REGION Network 18: MUTE 2
   RUNG wire#powerrail
      #Mute_LG_2_DB("I_S_Time_extension (TE)" := wire#w1, I_S_Material_selection_1 := wire#w2, "########## BASIC_INPUTS ##########" :=, I_S_ESPE_Channel_1 := #Light_Guard_Tuned, I_S_ESPE_Channel_2 := #Light_Guard_Tuned, "I_S_PLC_request (MR)" := #MR_2, I_S_Reset := #ACK, "I_S_Override hold-to-run-device" := #Bypass."Light Guards CX201 - CH1", I_S_first_logic_cycle := "FirstScan", I_S_Disc_Time_MR_and_TE :=, "########## MATERIAL_SELECTION_INPUTS ##########" :=, I_S_Material_selection_2 := #Material_Selection_2, I_S_Material_selection_3 :=, I_S_Material_selection_4 :=, "########## MATERIAL_TOLERANCE_LENGTH in mm ##########" :=, "I_S_Material_tolerance_length_Material_1-4" :=, "########## MAX_DISTANCE_MATERIAL_ESPE in mm ##########" :=, I_S_Max_distance_Material_to_ESPE := 200, "########## MATERIAL_LENGH_1-4 in mm ##########" :=, I_S_Material_length_Material_1 := 1000, I_S_Material_length_Material_2 := 800, I_S_Material_length_Material_3 :=, I_S_Material_length_Material_4 :=, "########## MATERIAL_SPEED_1-4 in mm/s ##########" :=, I_S_Material_speed_Material_1 := 167, I_S_Material_speed_Material_2 := 167, I_S_Material_speed_Material_3 :=, I_S_Material_speed_Material_4 :=, "########## BASIC_OUTPUTS ##########" =>, Q_Safety_release_1 =>, Q_Safety_release_2 =>, Q_SEE_Status =>, Q_Override_Status =>, Q_Reset_required =>, Q_Sequence_OK =>, "########## ERRORS ##########" =>, Error =>)
   END_RUNG
   RUNG wire#powerrail
      I_Contact( #MR_2 )
   END_RUNG wire#w1
   RUNG wire#powerrail
      I_Contact( #Material_Selection_2 )
   END_RUNG wire#w2
   // the same network as SCL:
   #Mute_LG_2_DB(I_S_ESPE_Channel_1 := #Light_Guard_Tuned,   // "SICK Safe Entry Exit HW PLC V02"
                 I_S_ESPE_Channel_2 := #Light_Guard_Tuned,
                 "I_S_PLC_request (MR)" := #MR_2,
                 "I_S_Time_extension (TE)" := NOT #MR_2,
                 I_S_Reset := #ACK,
                 "I_S_Override hold-to-run-device" := #Bypass."Light Guards CX201 - CH1",
                 I_S_first_logic_cycle := "FirstScan",
                 I_S_Material_selection_1 := NOT #Material_Selection_2,
                 I_S_Material_selection_2 := #Material_Selection_2,
                 I_S_Max_distance_Material_to_ESPE := 200,
                 I_S_Material_length_Material_1 := 1000,
                 I_S_Material_length_Material_2 := 800,
                 I_S_Material_speed_Material_1 := 167,
                 I_S_Material_speed_Material_2 := 167);
END_REGION

REGION Network 19: Gate 1 Sensor
   RUNG wire#powerrail
      #Gate_1_DB.ESTOP1(E_STOP := wire#w1, ACK_NEC :=, ACK := #ACK, TIME_DEL :=, Q =>, Q_DELAY =>, ACK_REQ =>, DIAG =>)
   END_RUNG
   RUNG wire#powerrail
      Contact( #Gate_1 )
   END_RUNG wire#w1
   RUNG wire#powerrail
      Contact( #Bypass.Gate_1 )
   END_RUNG wire#w1
   // the same network as SCL:
   #Gate_1_DB(E_STOP := #Gate_1 OR #Bypass.Gate_1, ACK := #ACK);   // ESTOP1
END_REGION

REGION Network 20: Gate 2 Sensor
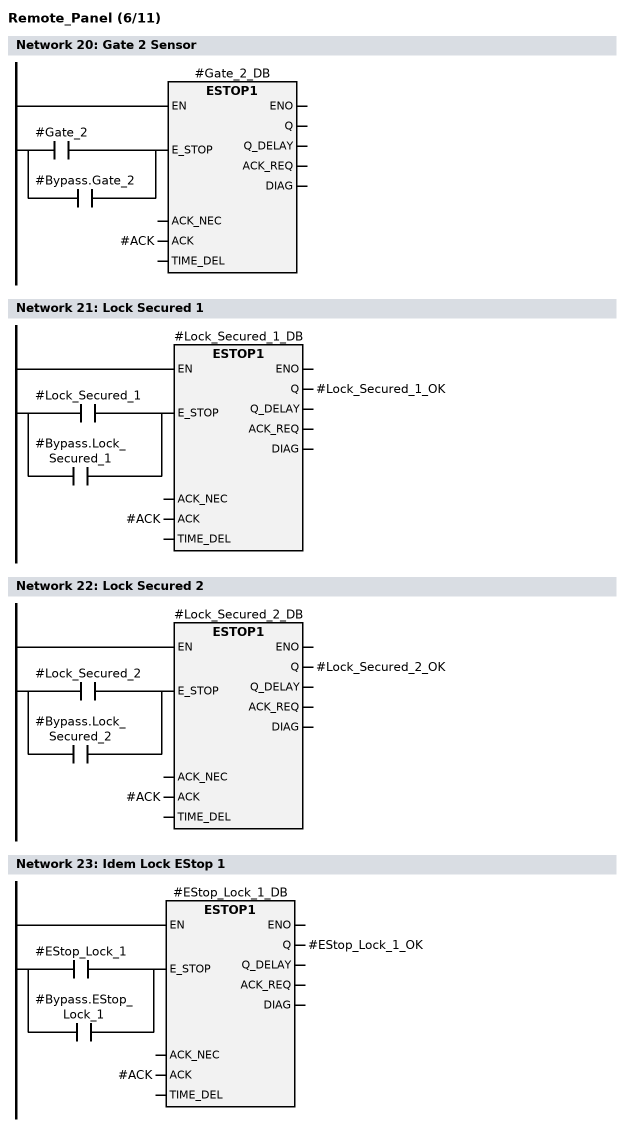
   RUNG wire#powerrail
      #Gate_2_DB.ESTOP1(E_STOP := wire#w1, ACK_NEC :=, ACK := #ACK, TIME_DEL :=, Q =>, Q_DELAY =>, ACK_REQ =>, DIAG =>)
   END_RUNG
   RUNG wire#powerrail
      Contact( #Gate_2 )
   END_RUNG wire#w1
   RUNG wire#powerrail
      Contact( #Bypass.Gate_2 )
   END_RUNG wire#w1
   // the same network as SCL:
   #Gate_2_DB(E_STOP := #Gate_2 OR #Bypass.Gate_2, ACK := #ACK);   // ESTOP1
END_REGION

REGION Network 21: Lock Secured 1
   RUNG wire#powerrail
      #Lock_Secured_1_DB.ESTOP1(E_STOP := wire#w1, ACK_NEC :=, ACK := #ACK, TIME_DEL :=, Q => #Lock_Secured_1_OK, Q_DELAY =>, ACK_REQ =>, DIAG =>)
   END_RUNG
   RUNG wire#powerrail
      Contact( #Lock_Secured_1 )
   END_RUNG wire#w1
   RUNG wire#powerrail
      Contact( #Bypass.Lock_Secured_1 )
   END_RUNG wire#w1
   // the same network as SCL:
   #Lock_Secured_1_DB(E_STOP := #Lock_Secured_1 OR #Bypass.Lock_Secured_1, ACK := #ACK, Q => #Lock_Secured_1_OK);   // ESTOP1
END_REGION

REGION Network 22: Lock Secured 2
   RUNG wire#powerrail
      #Lock_Secured_2_DB.ESTOP1(E_STOP := wire#w1, ACK_NEC :=, ACK := #ACK, TIME_DEL :=, Q => #Lock_Secured_2_OK, Q_DELAY =>, ACK_REQ =>, DIAG =>)
   END_RUNG
   RUNG wire#powerrail
      Contact( #Lock_Secured_2 )
   END_RUNG wire#w1
   RUNG wire#powerrail
      Contact( #Bypass.Lock_Secured_2 )
   END_RUNG wire#w1
   // the same network as SCL:
   #Lock_Secured_2_DB(E_STOP := #Lock_Secured_2 OR #Bypass.Lock_Secured_2, ACK := #ACK, Q => #Lock_Secured_2_OK);   // ESTOP1
END_REGION

REGION Network 23: Idem Lock EStop 1
   RUNG wire#powerrail
      #EStop_Lock_1_DB.ESTOP1(E_STOP := wire#w1, ACK_NEC :=, ACK := #ACK, TIME_DEL :=, Q => #EStop_Lock_1_OK, Q_DELAY =>, ACK_REQ =>, DIAG =>)
   END_RUNG
   RUNG wire#powerrail
      Contact( #EStop_Lock_1 )
   END_RUNG wire#w1
   RUNG wire#powerrail
      Contact( #Bypass.EStop_Lock_1 )
   END_RUNG wire#w1
   // the same network as SCL:
   #EStop_Lock_1_DB(E_STOP := #EStop_Lock_1 OR #Bypass.EStop_Lock_1, ACK := #ACK, Q => #EStop_Lock_1_OK);   // ESTOP1
END_REGION

REGION Network 24: Idem Lock EStop 2
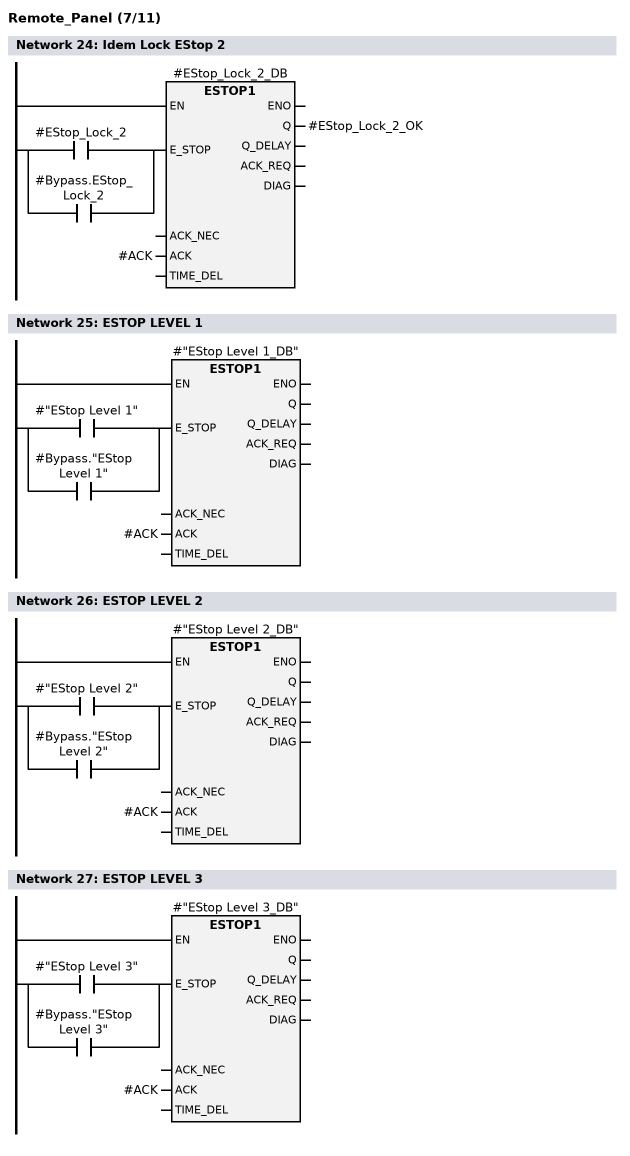
   RUNG wire#powerrail
      #EStop_Lock_2_DB.ESTOP1(E_STOP := wire#w1, ACK_NEC :=, ACK := #ACK, TIME_DEL :=, Q => #EStop_Lock_2_OK, Q_DELAY =>, ACK_REQ =>, DIAG =>)
   END_RUNG
   RUNG wire#powerrail
      Contact( #EStop_Lock_2 )
   END_RUNG wire#w1
   RUNG wire#powerrail
      Contact( #Bypass.EStop_Lock_2 )
   END_RUNG wire#w1
   // the same network as SCL:
   #EStop_Lock_2_DB(E_STOP := #EStop_Lock_2 OR #Bypass.EStop_Lock_2, ACK := #ACK, Q => #EStop_Lock_2_OK);   // ESTOP1
END_REGION

REGION Network 25: ESTOP LEVEL 1
   RUNG wire#powerrail
      #"EStop Level 1_DB".ESTOP1(E_STOP := wire#w1, ACK_NEC :=, ACK := #ACK, TIME_DEL :=, Q =>, Q_DELAY =>, ACK_REQ =>, DIAG =>)
   END_RUNG
   RUNG wire#powerrail
      Contact( #"EStop Level 1" )
   END_RUNG wire#w1
   RUNG wire#powerrail
      Contact( #Bypass."EStop Level 1" )
   END_RUNG wire#w1
   // the same network as SCL:
   #"EStop Level 1_DB"(E_STOP := #"EStop Level 1" OR #Bypass."EStop Level 1", ACK := #ACK);   // ESTOP1
END_REGION

REGION Network 26: ESTOP LEVEL 2
   RUNG wire#powerrail
      #"EStop Level 2_DB".ESTOP1(E_STOP := wire#w1, ACK_NEC :=, ACK := #ACK, TIME_DEL :=, Q =>, Q_DELAY =>, ACK_REQ =>, DIAG =>)
   END_RUNG
   RUNG wire#powerrail
      Contact( #"EStop Level 2" )
   END_RUNG wire#w1
   RUNG wire#powerrail
      Contact( #Bypass."EStop Level 2" )
   END_RUNG wire#w1
   // the same network as SCL:
   #"EStop Level 2_DB"(E_STOP := #"EStop Level 2" OR #Bypass."EStop Level 2", ACK := #ACK);   // ESTOP1
END_REGION

REGION Network 27: ESTOP LEVEL 3
   RUNG wire#powerrail
      #"EStop Level 3_DB".ESTOP1(E_STOP := wire#w1, ACK_NEC :=, ACK := #ACK, TIME_DEL :=, Q =>, Q_DELAY =>, ACK_REQ =>, DIAG =>)
   END_RUNG
   RUNG wire#powerrail
      Contact( #"EStop Level 3" )
   END_RUNG wire#w1
   RUNG wire#powerrail
      Contact( #Bypass."EStop Level 3" )
   END_RUNG wire#w1
   // the same network as SCL:
   #"EStop Level 3_DB"(E_STOP := #"EStop Level 3" OR #Bypass."EStop Level 3", ACK := #ACK);   // ESTOP1
END_REGION

REGION Network 28: ESTOP LEVEL 4
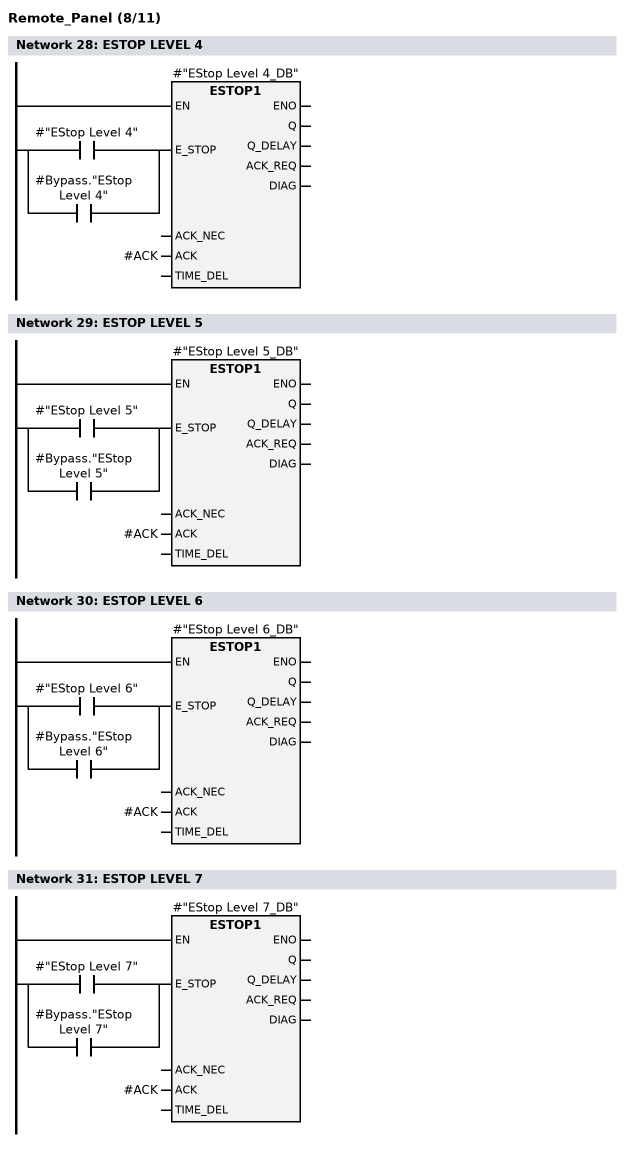
   RUNG wire#powerrail
      #"EStop Level 4_DB".ESTOP1(E_STOP := wire#w1, ACK_NEC :=, ACK := #ACK, TIME_DEL :=, Q =>, Q_DELAY =>, ACK_REQ =>, DIAG =>)
   END_RUNG
   RUNG wire#powerrail
      Contact( #"EStop Level 4" )
   END_RUNG wire#w1
   RUNG wire#powerrail
      Contact( #Bypass."EStop Level 4" )
   END_RUNG wire#w1
   // the same network as SCL:
   #"EStop Level 4_DB"(E_STOP := #"EStop Level 4" OR #Bypass."EStop Level 4", ACK := #ACK);   // ESTOP1
END_REGION

REGION Network 29: ESTOP LEVEL 5
   RUNG wire#powerrail
      #"EStop Level 5_DB".ESTOP1(E_STOP := wire#w1, ACK_NEC :=, ACK := #ACK, TIME_DEL :=, Q =>, Q_DELAY =>, ACK_REQ =>, DIAG =>)
   END_RUNG
   RUNG wire#powerrail
      Contact( #"EStop Level 5" )
   END_RUNG wire#w1
   RUNG wire#powerrail
      Contact( #Bypass."EStop Level 5" )
   END_RUNG wire#w1
   // the same network as SCL:
   #"EStop Level 5_DB"(E_STOP := #"EStop Level 5" OR #Bypass."EStop Level 5", ACK := #ACK);   // ESTOP1
END_REGION

REGION Network 30: ESTOP LEVEL 6
   RUNG wire#powerrail
      #"EStop Level 6_DB".ESTOP1(E_STOP := wire#w1, ACK_NEC :=, ACK := #ACK, TIME_DEL :=, Q =>, Q_DELAY =>, ACK_REQ =>, DIAG =>)
   END_RUNG
   RUNG wire#powerrail
      Contact( #"EStop Level 6" )
   END_RUNG wire#w1
   RUNG wire#powerrail
      Contact( #Bypass."EStop Level 6" )
   END_RUNG wire#w1
   // the same network as SCL:
   #"EStop Level 6_DB"(E_STOP := #"EStop Level 6" OR #Bypass."EStop Level 6", ACK := #ACK);   // ESTOP1
END_REGION

REGION Network 31: ESTOP LEVEL 7
   RUNG wire#powerrail
      #"EStop Level 7_DB".ESTOP1(E_STOP := wire#w1, ACK_NEC :=, ACK := #ACK, TIME_DEL :=, Q =>, Q_DELAY =>, ACK_REQ =>, DIAG =>)
   END_RUNG
   RUNG wire#powerrail
      Contact( #"EStop Level 7" )
   END_RUNG wire#w1
   RUNG wire#powerrail
      Contact( #Bypass."EStop Level 7" )
   END_RUNG wire#w1
   // the same network as SCL:
   #"EStop Level 7_DB"(E_STOP := #"EStop Level 7" OR #Bypass."EStop Level 7", ACK := #ACK);   // ESTOP1
END_REGION

REGION Network 32: ESTOP LEVEL 8
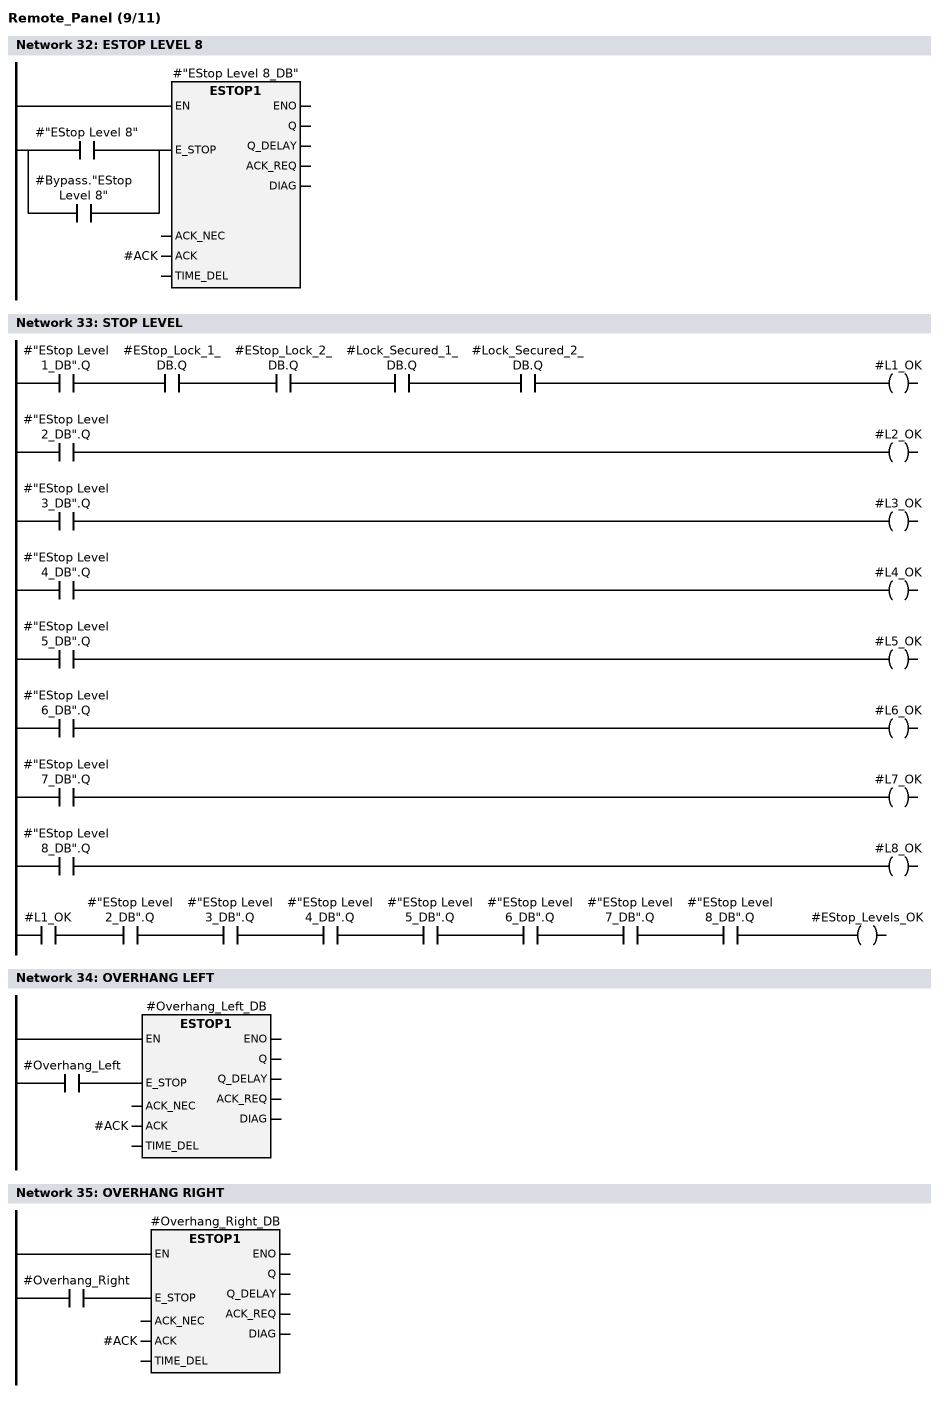
   RUNG wire#powerrail
      #"EStop Level 8_DB".ESTOP1(E_STOP := wire#w1, ACK_NEC :=, ACK := #ACK, TIME_DEL :=, Q =>, Q_DELAY =>, ACK_REQ =>, DIAG =>)
   END_RUNG
   RUNG wire#powerrail
      Contact( #"EStop Level 8" )
   END_RUNG wire#w1
   RUNG wire#powerrail
      Contact( #Bypass."EStop Level 8" )
   END_RUNG wire#w1
   // the same network as SCL:
   #"EStop Level 8_DB"(E_STOP := #"EStop Level 8" OR #Bypass."EStop Level 8", ACK := #ACK);   // ESTOP1
END_REGION

REGION Network 33: STOP LEVEL
   RUNG wire#powerrail
      Contact( #"EStop Level 1_DB".Q )
      Contact( #EStop_Lock_1_DB.Q )
      Contact( #EStop_Lock_2_DB.Q )
      Contact( #Lock_Secured_1_DB.Q )
      Contact( #Lock_Secured_2_DB.Q )
      Coil( #L1_OK )
   END_RUNG
   RUNG wire#powerrail
      Contact( #"EStop Level 2_DB".Q )
      Coil( #L2_OK )
   END_RUNG
   RUNG wire#powerrail
      Contact( #"EStop Level 3_DB".Q )
      Coil( #L3_OK )
   END_RUNG
   RUNG wire#powerrail
      Contact( #"EStop Level 4_DB".Q )
      Coil( #L4_OK )
   END_RUNG
   RUNG wire#powerrail
      Contact( #"EStop Level 5_DB".Q )
      Coil( #L5_OK )
   END_RUNG
   RUNG wire#powerrail
      Contact( #"EStop Level 6_DB".Q )
      Coil( #L6_OK )
   END_RUNG
   RUNG wire#powerrail
      Contact( #"EStop Level 7_DB".Q )
      Coil( #L7_OK )
   END_RUNG
   RUNG wire#powerrail
      Contact( #"EStop Level 8_DB".Q )
      Coil( #L8_OK )
   END_RUNG
   RUNG wire#powerrail
      Contact( #L1_OK )
      Contact( #"EStop Level 2_DB".Q )
      Contact( #"EStop Level 3_DB".Q )
      Contact( #"EStop Level 4_DB".Q )
      Contact( #"EStop Level 5_DB".Q )
      Contact( #"EStop Level 6_DB".Q )
      Contact( #"EStop Level 7_DB".Q )
      Contact( #"EStop Level 8_DB".Q )
      Coil( #EStop_Levels_OK )
   END_RUNG
   // the same network as SCL:
   #L1_OK := #"EStop Level 1_DB".Q AND #EStop_Lock_1_DB.Q AND #EStop_Lock_2_DB.Q AND #Lock_Secured_1_DB.Q AND #Lock_Secured_2_DB.Q;
   #L2_OK := #"EStop Level 2_DB".Q;
   #L3_OK := #"EStop Level 3_DB".Q;
   #L4_OK := #"EStop Level 4_DB".Q;
   #L5_OK := #"EStop Level 5_DB".Q;
   #L6_OK := #"EStop Level 6_DB".Q;
   #L7_OK := #"EStop Level 7_DB".Q;
   #L8_OK := #"EStop Level 8_DB".Q;
   #EStop_Levels_OK := #L1_OK AND #"EStop Level 2_DB".Q AND #"EStop Level 3_DB".Q AND #"EStop Level 4_DB".Q AND #"EStop Level 5_DB".Q AND #"EStop Level 6_DB".Q AND #"EStop Level 7_DB".Q AND #"EStop Level 8_DB".Q;
END_REGION

REGION Network 34: OVERHANG LEFT
   RUNG wire#powerrail
      #Overhang_Left_DB.ESTOP1(E_STOP := wire#w1, ACK_NEC :=, ACK := #ACK, TIME_DEL :=, Q =>, Q_DELAY =>, ACK_REQ =>, DIAG =>)
   END_RUNG
   RUNG wire#powerrail
      Contact( #Overhang_Left )
   END_RUNG wire#w1
   // the same network as SCL:
   #Overhang_Left_DB(E_STOP := #Overhang_Left, ACK := #ACK);   // ESTOP1
END_REGION

REGION Network 35: OVERHANG RIGHT
   RUNG wire#powerrail
      #Overhang_Right_DB.ESTOP1(E_STOP := wire#w1, ACK_NEC :=, ACK := #ACK, TIME_DEL :=, Q =>, Q_DELAY =>, ACK_REQ =>, DIAG =>)
   END_RUNG
   RUNG wire#powerrail
      Contact( #Overhang_Right )
   END_RUNG wire#w1
   // the same network as SCL:
   #Overhang_Right_DB(E_STOP := #Overhang_Right, ACK := #ACK);   // ESTOP1
END_REGION

REGION Network 36: Safety OK
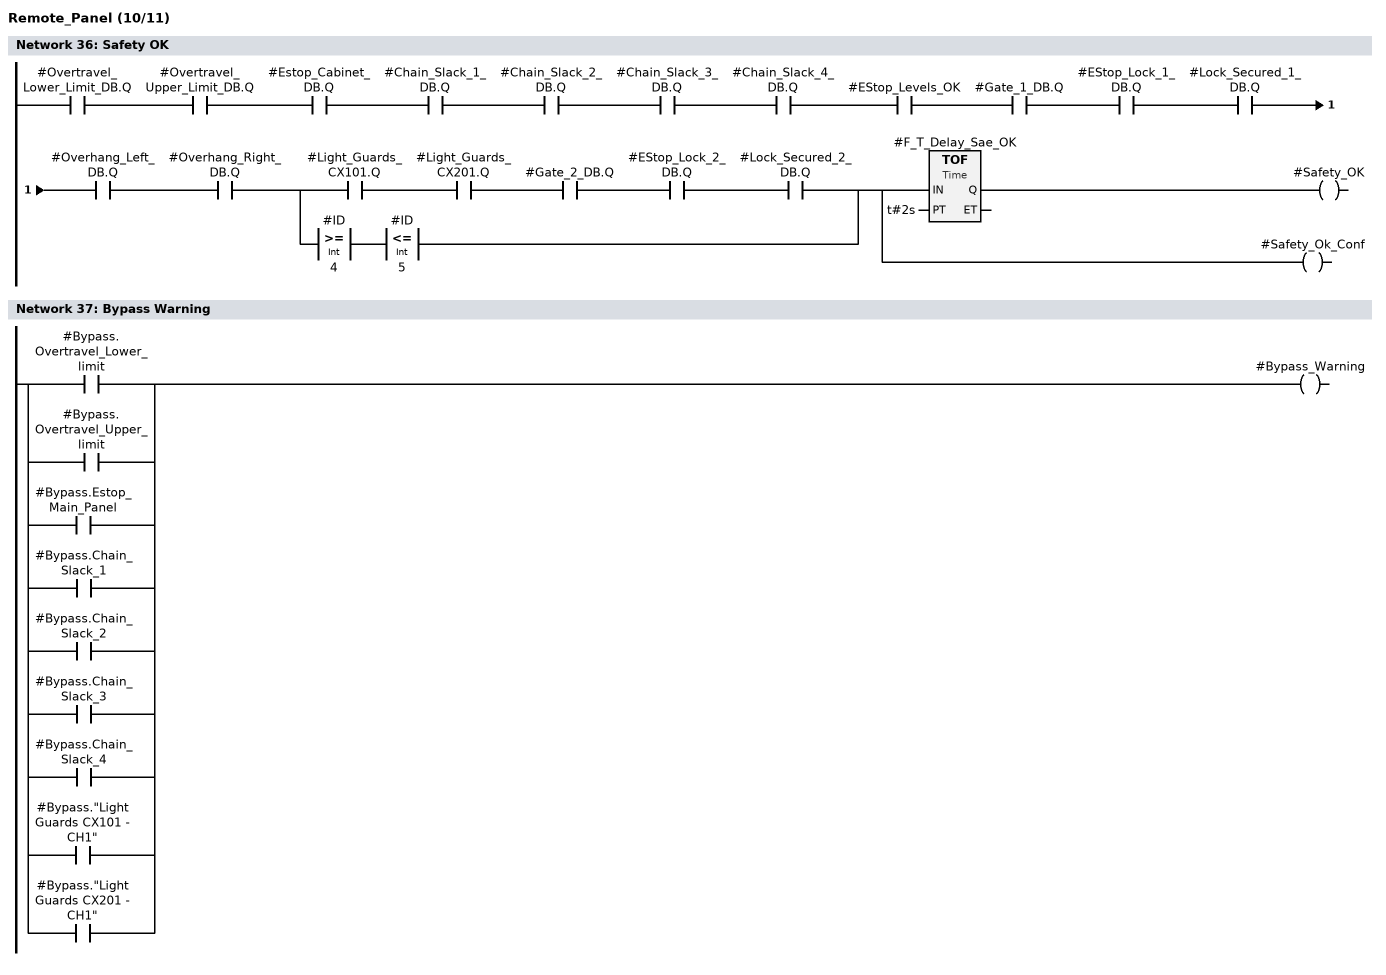
   RUNG wire#powerrail
      Contact( #Overtravel_Lower_Limit_DB.Q )
      Contact( #Overtravel_Upper_Limit_DB.Q )
      Contact( #Estop_Cabinet_DB.Q )
      Contact( #Chain_Slack_1_DB.Q )
      Contact( #Chain_Slack_2_DB.Q )
      Contact( #Chain_Slack_3_DB.Q )
      Contact( #Chain_Slack_4_DB.Q )
      Contact( #EStop_Levels_OK )
      Contact( #Gate_1_DB.Q )
      Contact( #EStop_Lock_1_DB.Q )
      Contact( #Lock_Secured_1_DB.Q )
      Contact( #Overhang_Left_DB.Q )
      Contact( #Overhang_Right_DB.Q )
      wire#w1
      Contact( #Light_Guards_CX101.Q )
      Contact( #Light_Guards_CX201.Q )
      Contact( #Gate_2_DB.Q )
      Contact( #EStop_Lock_2_DB.Q )
      Contact( #Lock_Secured_2_DB.Q )
      wire#w2
      { S7_Templates := "[time_type := Time, codedbool_type := DInt]" } #F_T_Delay_Sae_OK.TOF(pt := t#2s, et =>)
      Coil( #Safety_OK )
   END_RUNG
   RUNG wire#w1
      { S7_Templates := "SrcType := Int" } GE_Contact(in1 := #ID, in2 := 4)
      { S7_Templates := "SrcType := Int" } LE_Contact(in1 := #ID, in2 := 5)
   END_RUNG wire#w2
   RUNG wire#w2
      Coil( #Safety_Ok_Conf )
   END_RUNG
   // the same network as SCL:
   #_w1 := #Overtravel_Lower_Limit_DB.Q AND #Overtravel_Upper_Limit_DB.Q AND #Estop_Cabinet_DB.Q AND #Chain_Slack_1_DB.Q AND #Chain_Slack_2_DB.Q AND #Chain_Slack_3_DB.Q AND #Chain_Slack_4_DB.Q AND #EStop_Levels_OK AND #Gate_1_DB.Q AND #EStop_Lock_1_DB.Q AND #Lock_Secured_1_DB.Q AND #Overhang_Left_DB.Q AND #Overhang_Right_DB.Q AND ((#Light_Guards_CX101.Q AND #Light_Guards_CX201.Q AND #Gate_2_DB.Q AND #EStop_Lock_2_DB.Q AND #Lock_Secured_2_DB.Q) OR ((#ID >= 4) AND (#ID <= 5)));
   #F_T_Delay_Sae_OK.TOF(IN := #_w1, PT := t#2s);
   #Safety_OK := #F_T_Delay_Sae_OK.Q;
   #Safety_Ok_Conf := #_w1;
END_REGION

REGION Network 37: Bypass Warning
   RUNG wire#powerrail
      Contact( #Bypass.Overtravel_Lower_limit )
      wire#w1
      Coil( #Bypass_Warning )
   END_RUNG
   RUNG wire#powerrail
      Contact( #Bypass.Overtravel_Upper_limit )
   END_RUNG wire#w1
   RUNG wire#powerrail
      Contact( #Bypass.Estop_Main_Panel )
   END_RUNG wire#w1
   RUNG wire#powerrail
      Contact( #Bypass.Chain_Slack_1 )
   END_RUNG wire#w1
   RUNG wire#powerrail
      Contact( #Bypass.Chain_Slack_2 )
   END_RUNG wire#w1
   RUNG wire#powerrail
      Contact( #Bypass.Chain_Slack_3 )
   END_RUNG wire#w1
   RUNG wire#powerrail
      Contact( #Bypass.Chain_Slack_4 )
   END_RUNG wire#w1
   RUNG wire#powerrail
      Contact( #Bypass."Light Guards CX101 - CH1" )
   END_RUNG wire#w1
   RUNG wire#powerrail
      Contact( #Bypass."Light Guards CX201 - CH1" )
   END_RUNG wire#w1
   // the same network as SCL:
   #Bypass_Warning := #Bypass.Overtravel_Lower_limit OR #Bypass.Overtravel_Upper_limit OR #Bypass.Estop_Main_Panel OR #Bypass.Chain_Slack_1 OR #Bypass.Chain_Slack_2 OR #Bypass.Chain_Slack_3 OR #Bypass.Chain_Slack_4 OR #Bypass."Light Guards CX101 - CH1" OR #Bypass."Light Guards CX201 - CH1";
END_REGION

REGION Network 38: Enable outputs
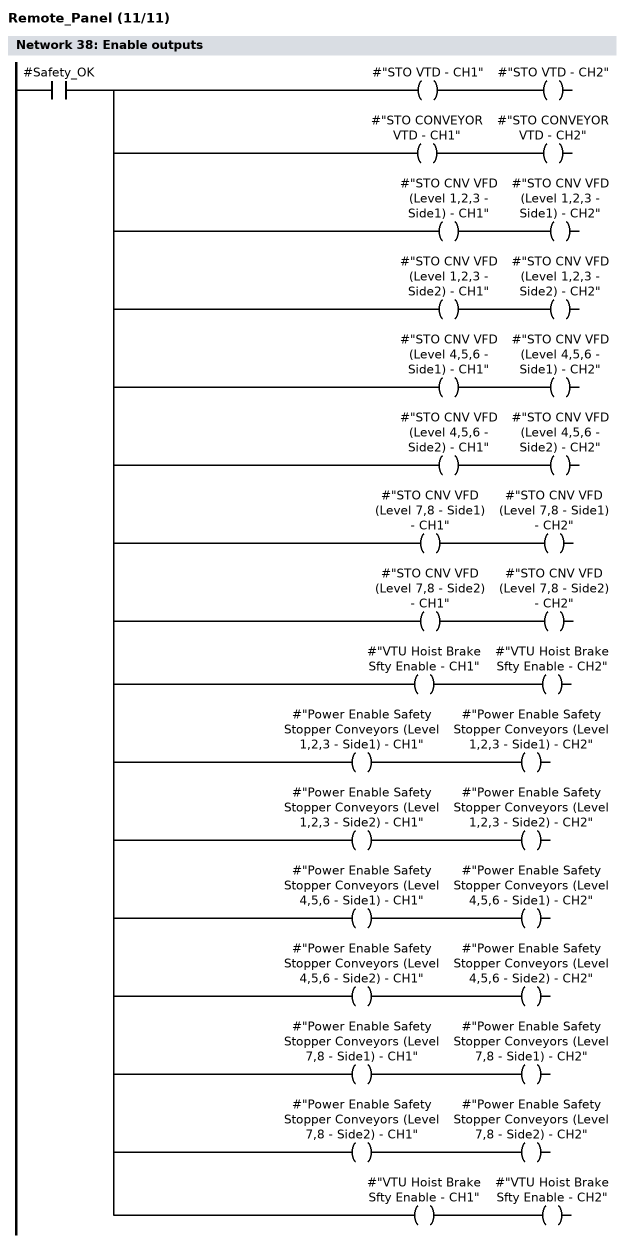
   RUNG wire#powerrail
      Contact( #Safety_OK )
      wire#w1
      Coil( #"STO VTD - CH1" )
      Coil( #"STO VTD - CH2" )
   END_RUNG
   RUNG wire#w1
      Coil( #"STO CONVEYOR VTD - CH1" )
      Coil( #"STO CONVEYOR VTD - CH2" )
   END_RUNG
   RUNG wire#w1
      Coil( #"STO CNV VFD (Level 1,2,3 - Side1) - CH1" )
      Coil( #"STO CNV VFD (Level 1,2,3 - Side1) - CH2" )
   END_RUNG
   RUNG wire#w1
      Coil( #"STO CNV VFD (Level 1,2,3 - Side2) - CH1" )
      Coil( #"STO CNV VFD (Level 1,2,3 - Side2) - CH2" )
   END_RUNG
   RUNG wire#w1
      Coil( #"STO CNV VFD (Level 4,5,6 - Side1) - CH1" )
      Coil( #"STO CNV VFD (Level 4,5,6 - Side1) - CH2" )
   END_RUNG
   RUNG wire#w1
      Coil( #"STO CNV VFD (Level 4,5,6 - Side2) - CH1" )
      Coil( #"STO CNV VFD (Level 4,5,6 - Side2) - CH2" )
   END_RUNG
   RUNG wire#w1
      Coil( #"STO CNV VFD (Level 7,8 - Side1) - CH1" )
      Coil( #"STO CNV VFD (Level 7,8 - Side1) - CH2" )
   END_RUNG
   RUNG wire#w1
      Coil( #"STO CNV VFD (Level 7,8 - Side2) - CH1" )
      Coil( #"STO CNV VFD (Level 7,8 - Side2) - CH2" )
   END_RUNG
   RUNG wire#w1
      Coil( #"VTU Hoist Brake Sfty Enable - CH1" )
      Coil( #"VTU Hoist Brake Sfty Enable - CH2" )
   END_RUNG
   RUNG wire#w1
      Coil( #"Power Enable Safety Stopper Conveyors (Level 1,2,3 - Side1) - CH1" )
      Coil( #"Power Enable Safety Stopper Conveyors (Level 1,2,3 - Side1) - CH2" )
   END_RUNG
   RUNG wire#w1
      Coil( #"Power Enable Safety Stopper Conveyors (Level 1,2,3 - Side2) - CH1" )
      Coil( #"Power Enable Safety Stopper Conveyors (Level 1,2,3 - Side2) - CH2" )
   END_RUNG
   RUNG wire#w1
      Coil( #"Power Enable Safety Stopper Conveyors (Level 4,5,6 - Side1) - CH1" )
      Coil( #"Power Enable Safety Stopper Conveyors (Level 4,5,6 - Side1) - CH2" )
   END_RUNG
   RUNG wire#w1
      Coil( #"Power Enable Safety Stopper Conveyors (Level 4,5,6 - Side2) - CH1" )
      Coil( #"Power Enable Safety Stopper Conveyors (Level 4,5,6 - Side2) - CH2" )
   END_RUNG
   RUNG wire#w1
      Coil( #"Power Enable Safety Stopper Conveyors (Level 7,8 - Side1) - CH1" )
      Coil( #"Power Enable Safety Stopper Conveyors (Level 7,8 - Side1) - CH2" )
   END_RUNG
   RUNG wire#w1
      Coil( #"Power Enable Safety Stopper Conveyors (Level 7,8 - Side2) - CH1" )
      Coil( #"Power Enable Safety Stopper Conveyors (Level 7,8 - Side2) - CH2" )
   END_RUNG
   RUNG wire#w1
      Coil( #"VTU Hoist Brake Sfty Enable - CH1" )
      Coil( #"VTU Hoist Brake Sfty Enable - CH2" )
   END_RUNG
   // the same network as SCL:
   #"STO VTD - CH1" := #Safety_OK;
   #"STO VTD - CH2" := #Safety_OK;
   #"STO CONVEYOR VTD - CH1" := #Safety_OK;
   #"STO CONVEYOR VTD - CH2" := #Safety_OK;
   #"STO CNV VFD (Level 1,2,3 - Side1) - CH1" := #Safety_OK;
   #"STO CNV VFD (Level 1,2,3 - Side1) - CH2" := #Safety_OK;
   #"STO CNV VFD (Level 1,2,3 - Side2) - CH1" := #Safety_OK;
   #"STO CNV VFD (Level 1,2,3 - Side2) - CH2" := #Safety_OK;
   #"STO CNV VFD (Level 4,5,6 - Side1) - CH1" := #Safety_OK;
   #"STO CNV VFD (Level 4,5,6 - Side1) - CH2" := #Safety_OK;
   #"STO CNV VFD (Level 4,5,6 - Side2) - CH1" := #Safety_OK;
   #"STO CNV VFD (Level 4,5,6 - Side2) - CH2" := #Safety_OK;
   #"STO CNV VFD (Level 7,8 - Side1) - CH1" := #Safety_OK;
   #"STO CNV VFD (Level 7,8 - Side1) - CH2" := #Safety_OK;
   #"STO CNV VFD (Level 7,8 - Side2) - CH1" := #Safety_OK;
   #"STO CNV VFD (Level 7,8 - Side2) - CH2" := #Safety_OK;
   #"VTU Hoist Brake Sfty Enable - CH1" := #Safety_OK;
   #"VTU Hoist Brake Sfty Enable - CH2" := #Safety_OK;
   #"Power Enable Safety Stopper Conveyors (Level 1,2,3 - Side1) - CH1" := #Safety_OK;
   #"Power Enable Safety Stopper Conveyors (Level 1,2,3 - Side1) - CH2" := #Safety_OK;
   #"Power Enable Safety Stopper Conveyors (Level 1,2,3 - Side2) - CH1" := #Safety_OK;
   #"Power Enable Safety Stopper Conveyors (Level 1,2,3 - Side2) - CH2" := #Safety_OK;
   #"Power Enable Safety Stopper Conveyors (Level 4,5,6 - Side1) - CH1" := #Safety_OK;
   #"Power Enable Safety Stopper Conveyors (Level 4,5,6 - Side1) - CH2" := #Safety_OK;
   #"Power Enable Safety Stopper Conveyors (Level 4,5,6 - Side2) - CH1" := #Safety_OK;
   #"Power Enable Safety Stopper Conveyors (Level 4,5,6 - Side2) - CH2" := #Safety_OK;
   #"Power Enable Safety Stopper Conveyors (Level 7,8 - Side1) - CH1" := #Safety_OK;
   #"Power Enable Safety Stopper Conveyors (Level 7,8 - Side1) - CH2" := #Safety_OK;
   #"Power Enable Safety Stopper Conveyors (Level 7,8 - Side2) - CH1" := #Safety_OK;
   #"Power Enable Safety Stopper Conveyors (Level 7,8 - Side2) - CH2" := #Safety_OK;
   #"VTU Hoist Brake Sfty Enable - CH1" := #Safety_OK;
   #"VTU Hoist Brake Sfty Enable - CH2" := #Safety_OK;
END_REGION
END_FUNCTION_BLOCK

FUNCTION_BLOCK "SICK Safe Entry Exit HW PLC V02"   // FB1000, F_FBD
TITLE = SICK Safe Entry Exit
AUTHOR : 2/29SD
FAMILY : S7-1500F
NAME : 9300351_02
VERSION : 2.0
// compiled for S7-1500F hardware controllers
// stored: IsIECCheckEnabled false, UDAEnableTagReadback false
   VAR_INPUT
      "########## BASIC_INPUTS ##########" : Bool := false;
      I_S_ESPE_Channel_1 : Bool := false;
      I_S_ESPE_Channel_2 : Bool := false;
      "I_S_PLC_request (MR)" : Bool := false;
      "I_S_Time_extension (TE)" : Bool := false;
      I_S_Reset : Bool := false;
      "I_S_Override hold-to-run-device" : Bool := false;
      I_S_first_logic_cycle : Bool := false;
      I_S_Disc_Time_MR_and_TE : Time := t#500ms;
      "########## MATERIAL_SELECTION_INPUTS ##########" : Bool := false;
      I_S_Material_selection_1 : Bool := false;
      I_S_Material_selection_2 : Bool := false;
      I_S_Material_selection_3 : Bool := false;
      I_S_Material_selection_4 : Bool := false;
      "########## MATERIAL_TOLERANCE_LENGTH in mm ##########" : Bool := false;
      "I_S_Material_tolerance_length_Material_1-4" : DInt := 100;
      "########## MAX_DISTANCE_MATERIAL_ESPE in mm ##########" : Bool := false;
      I_S_Max_distance_Material_to_ESPE : DInt := 0;
      "########## MATERIAL_LENGH_1-4 in mm ##########" : Bool := false;
      I_S_Material_length_Material_1 : DInt := 0;
      I_S_Material_length_Material_2 : DInt := 0;
      I_S_Material_length_Material_3 : DInt := 0;
      I_S_Material_length_Material_4 : DInt := 0;
      "########## MATERIAL_SPEED_1-4 in mm/s ##########" : Bool := false;
      I_S_Material_speed_Material_1 : DInt := 0;
      I_S_Material_speed_Material_2 : DInt := 0;
      I_S_Material_speed_Material_3 : DInt := 0;
      I_S_Material_speed_Material_4 : DInt := 0;
   END_VAR
   VAR_OUTPUT
      "########## BASIC_OUTPUTS ##########" : Bool := false;
      Q_Safety_release_1 : Bool := false;
      Q_Safety_release_2 : Bool;
      Q_SEE_Status : Bool := false;
      Q_Override_Status : Bool := false;
      Q_Reset_required : Bool := false;
      Q_Sequence_OK : Bool;
      "########## ERRORS ##########" : Bool := false;
      Error : Word := 0;
   END_VAR
   VAR
      "## BASIC SIGNALS ##" : Bool;
      ESPE : Bool;
      SEE_active : Bool;
      SEE_inactive : Bool;
      PLC_request : Bool;
      Time_extension : Bool;
      PLC_request_end : Bool;
      TE_signal_error : Bool;
      PLC_error : Bool;
      Timing_selection_error : Bool;
      Initiation_Error : Bool;
      SSE_aditional_release : Bool;
      Initiation : Bool;
      Termination : Bool;
      Termination_Seq_good : Bool;
      Override_status : Bool;
      Sequence_Signals_good : Bool;
      Material_1 : Bool;
      Material_2 : Bool;
      Material_3 : Bool;
      Material_4 : Bool;
      Min_time_good : Bool;
      Max_time_Error : Bool;
      TON_Tact_Lamps { S7_SetPoint := 'True'} : TON;
      TOF_Tact_Lamps { S7_SetPoint := 'True'} : TOF;
      Neg_Flag_Lamps : Bool;
      Blinking_tact : Bool;
      Always_0 : Bool := FALSE;
      Always_1 : Bool := TRUE;
      b_Sequence_Start : Bool;
      b_Sequence_OK : Bool;
      Sequence_OK { S7_SetPoint := 'True'} : TON;
      "## END BASIC SIGNALS ##" : Bool;
      "### CLOCK GENERATOR ###" : Bool;
      CLK_GEN_Edge_neg_1 : Bool;
      CLK_GEN_TON_Timer_1 { S7_SetPoint := 'True'} : TON;
      CLK_GEN_TOF_Timer_1 { S7_SetPoint := 'True'} : TOF;
      CLK_GEN_Tact : Bool;
      "### END CLOCK GENERATOR ###" : Bool;
      "### INITIATION ###" : Bool;
      INIT_HM_1 : Bool;
      INIT_HM_2 : Bool;
      INIT_HM_3 : Bool;
      INIT_Edge_neg_1 : Bool;
      "### END INITIATION ###" : Bool;
      "### MIN MAX TIME MONITORING ###" : Bool;
      MM_TIME_MONT_Fl_neg_1 : Bool;
      MM_TIME_MONT_TOF_Timer_1 { S7_SetPoint := 'True'} : TOF;
      MM_TIME_MONT_Int_timer_reset : Bool;
      MM_TIME_MONT_Counter_up_1 { S7_SetPoint := 'True'} : CTU;
      MM_TIME_MONT_Counter_up_2 { S7_SetPoint := 'True'} : CTU;
      MM_TIME_MONT_SEE_act_neg_edge : Bool;
      MM_TIME_MONT_Timer_reset : Bool;
      MM_TIME_MONT_TE_inactive : Bool;
      MM_TIME_MONT_TE_Timeout : Bool;
      MM_TIME_MONT_SEE_Timing_1 : Bool;
      MM_TIME_MONT_SEE_Timing_2 : Bool;
      MM_TIME_MONT_SEE_Timing_3 : Bool;
      MM_TIME_MONT_SEE_Timing_4 : Bool;
      "### END MIN MAX TIME MONITORING ###" : Bool;
      "### MULTIPLE STORE ###" : Bool;
      MUL_STORE_Edge_pos_1 : Bool;
      MUL_STORE_Save_Signal_1 : Bool;
      MUL_STORE_Save_Signal_2 : Bool;
      MUL_STORE_Save_Signal_3 : Bool;
      MUL_STORE_Save_Signal_4 : Bool;
      MUL_STORE_Save_Signal_5 : Bool;
      MUL_STORE_Save_Signal_6 : Bool;
      MUL_STORE_Save_Signal_7 : Bool;
      "### END MULTIPLE STORE ###" : Bool;
      "### OPERATION SELECTOR ###" : Bool;
      OP_SEL_Input_change : Bool;
      OP_SEL_Last_Cycle_Out_1 : Bool;
      OP_SEL_Last_Cycle_Out_2 : Bool;
      OP_SEL_Last_Cycle_Out_3 : Bool;
      OP_SEL_Last_Cycle_Out_4 : Bool;
      OP_SEL_Last_Cycle_Out_5 : Bool;
      OP_SEL_Last_Cycle_Out_6 : Bool;
      OP_SEL_Last_Cycle_Out_7 : Bool;
      OP_SEL_Last_Cycle_Out_8 : Bool;
      OP_SEL_HM_out_1 : Bool;
      OP_SEL_HM_out_2 : Bool;
      OP_SEL_HM_out_3 : Bool;
      OP_SEL_HM_out_4 : Bool;
      OP_SEL_HM_out_5 : Bool;
      OP_SEL_HM_out_6 : Bool;
      OP_SEL_HM_out_7 : Bool;
      OP_SEL_HM_out_8 : Bool;
      OP_SEL_TON_Timer_1 { S7_SetPoint := 'True'} : TON;
      OP_SEL_TON_Timer_2 { S7_SetPoint := 'True'} : TON;
      OP_SEL_Timing_1 : Bool;
      OP_SEL_Timing_2 : Bool;
      OP_SEL_Timing_3 : Bool;
      OP_SEL_Timing_4 : Bool;
      "### END OPERATION SELECTOR ###" : Bool;
      "### RESET1 ###" : Bool;
      RESET1_Edge_neg_1 : Bool;
      RESET1_M_Reset : Bool;
      RESET1_TON_TIMER_1 { S7_SetPoint := 'True'} : TON;
      RESET1_TON_TIMER_2 { S7_SetPoint := 'True'} : TON;
      RESET1_Release_OK : Bool;
      RESET1_Q : Bool;
      "### END RESET1 ###" : Bool;
      "### OVERRIDE ###" : Bool;
      OVR_TON_Timer_1 { S7_SetPoint := 'True'} : TON;
      OVR_Override_required : Bool;
      OVR_Override_status : Bool;
      OVR_Overriede_Clearance : Bool;
      "### END OVERRIDE ###" : Bool;
      "### RESET2 ###" : Bool;
      RESET2_Edge_neg_1 : Bool;
      RESET2_M_Reset : Bool;
      RESET2_TON_TIMER_1 { S7_SetPoint := 'True'} : TON;
      RESET2_TON_TIMER_2 { S7_SetPoint := 'True'} : TON;
      RESET2_Release_OK : Bool;
      "### END RESET2 ###" : Bool;
      "### TERMINATION ###" : Bool;
      TERM_Edge_neg_1 : Bool;
      TERM_Edge_pos_1 : Bool;
      TERM_HM_1 : Bool;
      TERM_TOF_Timer_1 { S7_SetPoint := 'True'} : TOF;
      "### END TERMINATION ###" : Bool;
      "### MIN_MAX_TIMER_RESET ###" : Bool;
      MIN_MAX_TIME_TON_Timer_Reset { S7_SetPoint := 'True'} : TON;
      "### END_MIN_MAX_TIMER_RESET ###" : Bool;
      "###MIN TIME  ###" : Bool;
      MIN_TIME_1_Timer_save : Time;
      MIN_TIME_1_Timer_1st_stop : Bool := FALSE;
      MIN_TIME_1_Edge_neg_1 : Bool;
      MIN_TIME_1_TON_Timer_1 { S7_SetPoint := 'True'} : TON;
      MIN_TIME_1_Q : Bool;
      MIN_TIME_2_Timer_save : Time;
      MIN_TIME_2_Timer_1st_stop : Bool := FALSE;
      MIN_TIME_2_Edge_neg : Bool;
      MIN_TIME_2_TON_Timer { S7_SetPoint := 'True'} : TON;
      MIN_TIME_2_Q : Bool;
      MIN_TIME_3_Timer_save : Time;
      MIN_TIME_3_Timer_1st_stop : Bool;
      MIN_TIME_3_Edge_neg : Bool;
      MIN_TIME_3_TON_Timer { S7_SetPoint := 'True'} : TON;
      MIN_TIME_3_Q : Bool;
      MIN_TIME_4_Timer_save : Time;
      MIN_TIME_4_Timer_1st_stop : Bool;
      MIN_TIME_4_Edge_neg : Bool;
      MIN_TIME_4_TON_Timer { S7_SetPoint := 'True'} : TON;
      MIN_TIME_4_Q : Bool;
      "###END MIN TIME ###" : Bool;
      "###MAX TIME  ###" : Bool;
      MAX_TIME_1_Timer_save : Time;
      MAX_TIME_1_Timer_1st_stop : Bool;
      MAX_TIME_1_Edge_neg : Bool;
      MAX_TIME_1_TON_Timer { S7_SetPoint := 'True'} : TON;
      MAX_TIME_1_Q : Bool;
      MAX_TIME_2_Timer_save : Time;
      MAX_TIME_2_Timer_1st_stop : Bool;
      MAX_TIME_2_Edge_neg : Bool;
      MAX_TIME_2_TON_Timer { S7_SetPoint := 'True'} : TON;
      MAX_TIME_2_Q : Bool;
      MAX_TIME_3_Timer_save : Time;
      MAX_TIME_3_Timer_1st_stop : Bool;
      MAX_TIME_3_Edge_neg : Bool;
      MAX_TIME_3_TON_Timer { S7_SetPoint := 'True'} : TON;
      MAX_TIME_3_Q : Bool;
      MAX_TIME_4_Timer_save : Time;
      MAX_TIME_4_Timer_1st_stop : Bool;
      MAX_TIME_4_Edge_neg : Bool;
      MAX_TIME_4_TON_Timer { S7_SetPoint := 'True'} : TON;
      MAX_TIME_4_Q : Bool;
      "###END MAX TIME  ###" : Bool;
      "### DISC CONTROL 1 ###" : Bool;
      DISC_1_b_Input_A : Bool;
      DISC_1_b_Input_B : Bool;
      DISC_1_Fl_pos_1 : Bool;
      DISC_1_Fl_neg_1 : Bool;
      DISC_1_Fl_neg_2 : Bool;
      DISC_1_Startbit : Bool;
      DISC_1_Stopbit : Bool;
      DISC_1_M_Release : Bool;
      DISC_1_M_AND_Mode_active : Bool;
      DISC_1_TON_Timer_1 { S7_SetPoint := 'True'} : TON;
      DISC_1_TON_Timer_2 { S7_SetPoint := 'True'} : TON;
      DISC_1_TON_Timer_3 { S7_SetPoint := 'True'} : TON;
      DISC_1_TOF_Timer_1 { S7_SetPoint := 'True'} : TOF;
      DISC_1_TOF_Timer_2 { S7_SetPoint := 'True'} : TOF;
      DISC_1_Q : Bool;
      DISC_1_Error : Bool;
      DISC_1_Error_Discrepancy_1 : Bool;
      DISC_1_Error_Discrepancy_2 : Bool;
      "### END DISC CONTROL 1 ###" : Bool;
      "### DISC CONTROL 2 ###" : Bool;
      DISC_2_b_Input_A : Bool;
      DISC_2_b_Input_B : Bool;
      DISC_2_Fl_pos_1 : Bool;
      DISC_2_Fl_neg_1 : Bool;
      DISC_2_Fl_neg_2 : Bool;
      DISC_2_Startbit : Bool;
      DISC_2_Stopbit : Bool;
      DISC_2_M_Release : Bool;
      DISC_2_M_AND_Mode_active : Bool;
      DISC_2_TON_Timer_1 { S7_SetPoint := 'True'} : TON;
      DISC_2_TON_Timer_2 { S7_SetPoint := 'True'} : TON;
      DISC_2_TON_Timer_3 { S7_SetPoint := 'True'} : TON;
      DISC_2_TOF_Timer_1 { S7_SetPoint := 'True'} : TOF;
      DISC_2_TOF_Timer_2 { S7_SetPoint := 'True'} : TOF;
      DISC_2_Q : Bool;
      DISC_2_Error : Bool;
      DISC_2_Error_Discrepancy_2 : Bool;
      DISC_2_Error_Discrepancy_1 : Bool;
      "### END DISC CONTROL 2 ###" : Bool;
      "### PLC SIG MONITORING ###" : Bool;
      PLC_SIG_MON_Edge_pos_1 : Bool;
      PLC_SIG_MON_Edge_neg_1 : Bool;
      PLC_SIG_MON_Edge_neg_2 : Bool;
      PLC_SIG_MON_HM_1 : Bool;
      PLC_SIG_MON_Int_muting_request : Bool;
      PLC_SIG_MON_Int_time_extension : Bool;
      PLC_SIG_MON_Discrepancy_control_Q : Bool;
      PLC_SIG_MON_Error_discrepancy_control_1 : Bool;
      PLC_SIG_MON_TON_Timer_1 { S7_SetPoint := 'True'} : TON;
      "### END PLC SIG MONITORING ###" : Bool;
      "### SSE #####" : Bool;
      SSE_Int_Enable : Bool;
      SSE_Int_Muting_active : Bool;
      SSE_Int_Safe_condition : Bool;
      "### END SSE #####" : Bool;
      "### SEQUENCE MONITORING ###" : Bool;
      SEQ_MON_TOF_Timer_1 { S7_SetPoint := 'True'} : TOF;
      SEQ_MON_TOF_Timer_2 { S7_SetPoint := 'True'} : TOF;
      SEQ_MON_TOF_Timer_3 { S7_SetPoint := 'True'} : TOF;
      SEQ_MON_TOF_Timer_4 { S7_SetPoint := 'True'} : TOF;
      SEQ_MON_TON_Timer_5 { S7_SetPoint := 'True'} : TON;
      SEQ_MON_TON_Timer_6 { S7_SetPoint := 'True'} : TON;
      SEQ_MON_TON_Timer_7 { S7_SetPoint := 'True'} : TON;
      SEQ_MON_TON_Timer_8 { S7_SetPoint := 'True'} : TON;
      SEQ_MON_TON_Timer_9 { S7_SetPoint := 'True'} : TON;
      SEQ_MON_TON_Timer_10 { S7_SetPoint := 'True'} : TON;
      SEQ_MON_TON_Timer_11 { S7_SetPoint := 'True'} : TON;
      SEQ_MON_TON_Timer_12 { S7_SetPoint := 'True'} : TON;
      SEQ_MON_Edge_PLC_request : Bool;
      SEQ_MON_Edge_pos_1 : Bool;
      SEQ_MON_Error_PLC_Req : Bool;
      SEQ_MON_HM_PLC_request : Bool;
      "### END SEQUENCE MONITORING ###" : Bool;
      "### ERROR HANDLING ###" : Bool;
      ERR_Handling_INT : Int;
      ERR_Handling_Neg_Flag : Bool;
      ERR_Signal_monitoring_MR_TE : Bool;
      ERR_Signal_monitoring_MR_TE_direct : Bool;
      HM_Sequenz_MR_TE_1 : Bool;
      HM_Sequenz_MR_TE_2 : Bool;
      HM_Sequenz_MR_TE_OK : Bool;
      ERR_Flag_Pos : Bool;
      ERR_FL_Neg : Bool;
      TON_Timer_Err_direct { S7_SetPoint := 'True'} : TON;
      "Create Error Termination Sequence" : Bool;
      "Create Error Min time" : Bool;
      "Create Error Max time" : Bool;
      "Create Error Timing selection" : Bool;
      "Create Error PLC Signal" : Bool;
      "Create Error TE Signal" : Bool;
      "Create Error Discrepancy MR TE" : Bool;
      "Create Error Discrepancy ESPE" : Bool;
      "Create Error calculation zero" : Bool;
      "Create Error Signal monitoring MR TE" : Bool;
      "Create Error Max. Dist ESPE" : Bool;
      "Create Error Monitoring Max. Muting" : Bool;
      "Create Error Max. INIT Time" : Bool;
      "Create Error Initiation sequence" : Bool;
      "Create Error min time less 500mm" : Bool;
      Reset_bit : Bool;
      "### END ERROR HANDLING ###" : Bool;
   END_VAR
BEGIN
END_FUNCTION_BLOCK

FUNCTION "Overhang_IO_FC" : Void   // FC40, F_LAD
{ S7_Optimized_Access := 'TRUE' }
VERSION : 0.1
// stored: AutoNumber true, IsIECCheckEnabled false, UDAEnableTagReadback false
BEGIN

REGION Network 1: SYSTEM 1
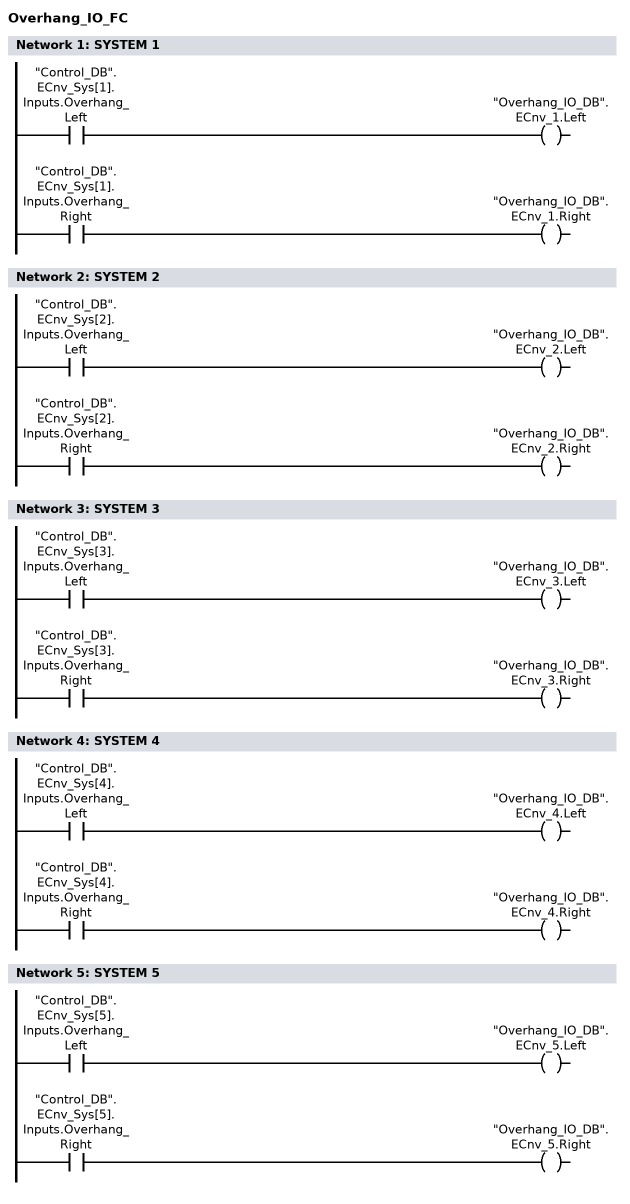
   RUNG wire#powerrail
      Contact( "Control_DB".ECnv_Sys[1].Inputs.Overhang_Left )
      Coil( "Overhang_IO_DB".ECnv_1.Left )
   END_RUNG
   RUNG wire#powerrail
      Contact( "Control_DB".ECnv_Sys[1].Inputs.Overhang_Right )
      Coil( "Overhang_IO_DB".ECnv_1.Right )
   END_RUNG
   // the same network as SCL:
   "Overhang_IO_DB".ECnv_1.Left := "Control_DB".ECnv_Sys[1].Inputs.Overhang_Left;
   "Overhang_IO_DB".ECnv_1.Right := "Control_DB".ECnv_Sys[1].Inputs.Overhang_Right;
END_REGION

REGION Network 2: SYSTEM 2
   RUNG wire#powerrail
      Contact( "Control_DB".ECnv_Sys[2].Inputs.Overhang_Left )
      Coil( "Overhang_IO_DB".ECnv_2.Left )
   END_RUNG
   RUNG wire#powerrail
      Contact( "Control_DB".ECnv_Sys[2].Inputs.Overhang_Right )
      Coil( "Overhang_IO_DB".ECnv_2.Right )
   END_RUNG
   // the same network as SCL:
   "Overhang_IO_DB".ECnv_2.Left := "Control_DB".ECnv_Sys[2].Inputs.Overhang_Left;
   "Overhang_IO_DB".ECnv_2.Right := "Control_DB".ECnv_Sys[2].Inputs.Overhang_Right;
END_REGION

REGION Network 3: SYSTEM 3
   RUNG wire#powerrail
      Contact( "Control_DB".ECnv_Sys[3].Inputs.Overhang_Left )
      Coil( "Overhang_IO_DB".ECnv_3.Left )
   END_RUNG
   RUNG wire#powerrail
      Contact( "Control_DB".ECnv_Sys[3].Inputs.Overhang_Right )
      Coil( "Overhang_IO_DB".ECnv_3.Right )
   END_RUNG
   // the same network as SCL:
   "Overhang_IO_DB".ECnv_3.Left := "Control_DB".ECnv_Sys[3].Inputs.Overhang_Left;
   "Overhang_IO_DB".ECnv_3.Right := "Control_DB".ECnv_Sys[3].Inputs.Overhang_Right;
END_REGION

REGION Network 4: SYSTEM 4
   RUNG wire#powerrail
      Contact( "Control_DB".ECnv_Sys[4].Inputs.Overhang_Left )
      Coil( "Overhang_IO_DB".ECnv_4.Left )
   END_RUNG
   RUNG wire#powerrail
      Contact( "Control_DB".ECnv_Sys[4].Inputs.Overhang_Right )
      Coil( "Overhang_IO_DB".ECnv_4.Right )
   END_RUNG
   // the same network as SCL:
   "Overhang_IO_DB".ECnv_4.Left := "Control_DB".ECnv_Sys[4].Inputs.Overhang_Left;
   "Overhang_IO_DB".ECnv_4.Right := "Control_DB".ECnv_Sys[4].Inputs.Overhang_Right;
END_REGION

REGION Network 5: SYSTEM 5
   RUNG wire#powerrail
      Contact( "Control_DB".ECnv_Sys[5].Inputs.Overhang_Left )
      Coil( "Overhang_IO_DB".ECnv_5.Left )
   END_RUNG
   RUNG wire#powerrail
      Contact( "Control_DB".ECnv_Sys[5].Inputs.Overhang_Right )
      Coil( "Overhang_IO_DB".ECnv_5.Right )
   END_RUNG
   // the same network as SCL:
   "Overhang_IO_DB".ECnv_5.Left := "Control_DB".ECnv_Sys[5].Inputs.Overhang_Left;
   "Overhang_IO_DB".ECnv_5.Right := "Control_DB".ECnv_Sys[5].Inputs.Overhang_Right;
END_REGION
END_FUNCTION

FUNCTION "Mode_Change_F" : Void   // FC2, SCL
{ S7_Optimized_Access := 'TRUE' }
VERSION : 0.1
// stored: AutoNumber true, IsIECCheckEnabled false, SetENOAutomatically false, UDAEnableTagReadback false
   VAR_INPUT
      Mode : UInt;
   END_VAR
   VAR_TEMP
      i : UInt;
      j : UInt;
   END_VAR
BEGIN
   // REGION Change all devices
   //     "Control_DB".ECnv_Control.Instruction.Mode_Change := #Mode;
   //     "Control_DB".VTD_Control.Instruction.Mode_Change := #Mode;

   //     FOR #i := "Settings_DB".VTD_Settings.Lowest_Level TO "Settings_DB".VTD_Settings.Highest_Level DO
   //         "Control_DB".LCnv_Control.Cnv_Level_Control[#i].Cnv1_Control.Instruction.Mode_Change := #Mode;
   //         "Control_DB".LCnv_Control.Cnv_Level_Control[#i].Cnv2_Control.Instruction.Mode_Change := #Mode;
   //     END_FOR;
   // END_REGION
END_FUNCTION

FUNCTION "OT_Charge_Commands" : Void   // FC52, SCL
{ S7_Optimized_Access := 'TRUE' }
VERSION : 0.1
// stored: AutoNumber true, IsIECCheckEnabled false, SetENOAutomatically false, UDAEnableTagReadback false
   VAR_IN_OUT
      Auto_Test : "Auto_Test";
   END_VAR
BEGIN
   "OrderTable_HMI"."Manual order" := #Auto_Test.Manual;
   //PALLET TYPE
   IF #Auto_Test."Pallet Type" = 'C' THEN
       "OrderTable_HMI"."Pallet Type" := 1;
   ELSIF #Auto_Test."Pallet Type" = 'E' THEN
       "OrderTable_HMI"."Pallet Type" := 2;
   END_IF;
   //TOWER 1 PALLET ALIGNMENT
   IF #Auto_Test."Tower 1 Pallet Alignment" = 'R' THEN
       "OrderTable_HMI"."Tower 1 Pallet Alignment" := 1;
   ELSIF #Auto_Test."Tower 1 Pallet Alignment" = 'L' THEN
       "OrderTable_HMI"."Tower 1 Pallet Alignment" := 2;
   END_IF;
   //TOWER 2 PALLET ALIGNMENT
   IF #Auto_Test."Tower 2 Pallet Alignment" = 'R' THEN
       "OrderTable_HMI"."Tower 2 Pallet Alignment" := 1;
   ELSIF #Auto_Test."Tower 2 Pallet Alignment" = 'L' THEN
       "OrderTable_HMI"."Tower 2 Pallet Alignment" := 2;
   END_IF;
   //ECONVEYOR PALLET ALIGNMENT
   IF #Auto_Test."Extractor Pallet Alignment" = 'R' THEN
       "OrderTable_HMI"."Extractor Pallet Alignment" := 1;
   ELSIF #Auto_Test."Extractor Pallet Alignment" = 'L' THEN
       "OrderTable_HMI"."Extractor Pallet Alignment" := 2;
   ELSIF #Auto_Test."Extractor Pallet Alignment" = 'C' THEN
       "OrderTable_HMI"."Extractor Pallet Alignment" := 3;
   END_IF;
   "OrderTable_HMI"."From level" := #Auto_Test."From level";
   "OrderTable_HMI"."To level" := #Auto_Test."To level";
   "OrderTable_HMI"."Testing Time" := #Auto_Test."Testing Time";
   "OrderTable_HMI"."Numer of cycles" := #Auto_Test."Numer of cycles";
   "OrderTable_HMI".Level := UINT_TO_BYTE(#Auto_Test.Level);
   "OrderTable_HMI".Tower := UINT_TO_BYTE(#Auto_Test.Tower);
END_FUNCTION

FUNCTION "OT_Charge_Commands_1" : Void   // FC64, SCL
{ S7_Optimized_Access := 'TRUE' }
VERSION : 0.1
// stored: AutoNumber true, IsIECCheckEnabled false, SetENOAutomatically false, UDAEnableTagReadback false
   VAR_IN_OUT
      Auto_Test : "Auto_Test_1";
   END_VAR
BEGIN
   "OrderTable_HMI"."Manual order" := #Auto_Test.Manual;
   //PALLET TYPE
   IF #Auto_Test."Pallet Type" = 'C' THEN
       "OrderTable_HMI"."Pallet Type" := 1;
   ELSIF #Auto_Test."Pallet Type" = 'E' THEN
       "OrderTable_HMI"."Pallet Type" := 2;
   END_IF;
   //TOWER 1 PALLET ALIGNMENT
   IF #Auto_Test."Tower 1 Pallet Alignment" = 'R' THEN
       "OrderTable_HMI"."Tower 1 Pallet Alignment" := 1;
   ELSIF #Auto_Test."Tower 1 Pallet Alignment" = 'L' THEN
       "OrderTable_HMI"."Tower 1 Pallet Alignment" := 2;
   END_IF;
   //ECONVEYOR PALLET ALIGNMENT
   IF #Auto_Test."Extractor Pallet Alignment" = 'R' THEN
       "OrderTable_HMI"."Extractor Pallet Alignment" := 1;
   ELSIF #Auto_Test."Extractor Pallet Alignment" = 'L' THEN
       "OrderTable_HMI"."Extractor Pallet Alignment" := 2;
   ELSIF #Auto_Test."Extractor Pallet Alignment" = 'C' THEN
       "OrderTable_HMI"."Extractor Pallet Alignment" := 3;
   END_IF;
   "OrderTable_HMI"."From level" := #Auto_Test."From level";
   "OrderTable_HMI"."To level" := #Auto_Test."To level";
   "OrderTable_HMI"."Testing Time" := #Auto_Test."Testing Time";
   "OrderTable_HMI"."Numer of cycles" := #Auto_Test."Numer of cycles";
   "OrderTable_HMI".Level := UINT_TO_BYTE(#Auto_Test.Level);
   "OrderTable_HMI".Tower := UINT_TO_BYTE(#Auto_Test.Tower);
END_FUNCTION

FUNCTION "ParseShuttle_Status" : "Shuttle_MQTT_Status_Msg"   // FC16, SCL
{ S7_Optimized_Access := 'TRUE' }
VERSION : 0.1
// stored: AutoNumber true, IsIECCheckEnabled false, SetENOAutomatically false, UDAEnableTagReadback false
   VAR_INPUT
      String_1 : String;
      String_2 : String;
      String_3 : String;
      String_4 : String;
      String_5 : String;
      String_6 : String;
   END_VAR
   VAR CONSTANT
      Empty : String;
   END_VAR
BEGIN
   #ParseShuttle_Status.Request_ID := "FindDINTFieldFragmented"(FieldName := 'requestId',
                                                                Str1 := #String_1,
                                                                Str2:=#Empty);
   #ParseShuttle_Status.Position_ID := "FindDINTFieldFragmented"(FieldName := 'positionId',
                                                                 Str1 := #String_1,
                                                                 Str2 := #Empty);
   #ParseShuttle_Status.Destination_ID := "FindDINTFieldFragmented"(FieldName := 'destinationId',
                                                                    Str1 := #String_1,
                                                                    Str2:=#Empty);
   #ParseShuttle_Status.Distance_Remaining := "FindDINTFieldFragmented"(FieldName := 'distanceRemaining',
                                                                        Str1 := #String_1,
                                                                        Str2 := #Empty);
   #ParseShuttle_Status.Position_X := "FindDINTFieldFragmented"(FieldName := 'positionX',
                                                                Str1 := #String_1,
                                                                Str2 := #Empty);
   #ParseShuttle_Status.Position_Y := "FindDINTFieldFragmented"(FieldName := 'positionY',
                                                                Str1 := #String_1,
                                                                Str2 := #Empty);
   #ParseShuttle_Status.Floor := "FindIntField"(FieldName := 'floor',
                                                   JsonStr := #String_1);
   #ParseShuttle_Status.Operation_Mode := "FindStringField"(FieldName := 'operationMode',
                                                            JsonStr := #String_1);
   #ParseShuttle_Status.Operational_State := "FindStringField"(FieldName := 'operationState',
                                                               JsonStr := #String_2);
   #ParseShuttle_Status.Load_State := "FindStringField"(FieldName := 'loadState',
                                                        JsonStr := #String_2);
   #ParseShuttle_Status.Error_Vehicle_1 := INT_TO_UINT("FindINTFieldFragmented"(FieldName := 'errorVehicle1',
                                                                                                                                    Str1 := #String_2,
                                                                                                                                    Str2:=#String_2));
   #ParseShuttle_Status.Error_Vehicle_2 := INT_TO_UINT("FindIntField"(FieldName := 'errorVehicle2',
                                                                                                                          JsonStr := #String_2));
   #ParseShuttle_Status.Error_Vehicle_3 := INT_TO_UINT("FindIntField"(FieldName := 'errorVehicle3',
                                                                                                                          JsonStr := #String_3));
   #ParseShuttle_Status.Error_Vehicle_4 := INT_TO_UINT("FindIntField"(FieldName := 'errorVehicle4',
                                                                                                                          JsonStr := #String_3));
   #ParseShuttle_Status.Error_Vehicle_5 := INT_TO_UINT("FindIntField"(FieldName := 'errorVehicle5',
                                                                                                                          JsonStr := #String_3));
   #ParseShuttle_Status.Error_Vehicle_6 := INT_TO_UINT("FindIntField"(FieldName := 'errorVehicle6',
                                                                                                                          JsonStr := #String_4));
   #ParseShuttle_Status.Sensor_Inputs := INT_TO_UINT("FindIntField"(FieldName := 'sensorInputs',
                                                                                                                      JsonStr := #String_4));
   #ParseShuttle_Status.Sensor_Outputs := INT_TO_UINT("FindIntField"(FieldName := 'sensorOutputs',
                                                                                                                        JsonStr := #String_4));
   #ParseShuttle_Status.Reader_Value := "FindDINTFieldFragmented"(FieldName := 'readerValue',
                                                                  Str1 := #String_4,
                                                                Str2 := #Empty);
   #ParseShuttle_Status.Pallet_Type := "FindStringField"(FieldName := 'palletType',
                                                         JsonStr := #String_4);
   #ParseShuttle_Status.Energy_Level := INT_TO_UINT("FindINTFieldFragmented"(FieldName := 'energyLevel',
                                                                                                                              Str1 := #String_5,
                                                                                                                              Str2:=#String_5));
   #ParseShuttle_Status.Battery_Voltage := INT_TO_UINT("FindIntField"(FieldName := 'batteryVoltage',
                                                                                                                          JsonStr := #String_5));
   #ParseShuttle_Status.Paused := "FindBoolField"(FieldName := 'paused',
                                                  JsonStr := #String_5);
   #ParseShuttle_Status.Last_Received_Order_ID := "FindIntField"(FieldName := 'lastReceivedOrderId',
                                                                 JsonStr := #String_5);
    #ParseShuttle_Status.Current_Order_ID := "FindIntField"(FieldName := 'currentOrderId',
                                                            JsonStr := #String_6);
          #ParseShuttle_Status.Last_Finished_Order_ID := "FindIntField"(FieldName := 'lastFinishedOrderId',
                                                                        JsonStr := #String_6);
END_FUNCTION

FUNCTION "PopUp_Screens" : Void   // FC9, SCL
{ S7_Optimized_Access := 'TRUE' }
VERSION : 0.1
// stored: AutoNumber true, IsIECCheckEnabled false, SetENOAutomatically false, UDAEnableTagReadback false
BEGIN
   //VTD SETTINGS
   IF "VTD_System_Selected_HMI" <> 0 (*AND "HMI_DB".ScreenNo_Main = 11*) AND "PopUps_DB".VTD_Settings.ID = "Settings_System_Selected" THEN
       CASE "Settings_System_Selected" OF
           1:
               "Settings_DB".VTD_Sys[1] := "PopUps_DB".VTD_Settings;
               "Settings_Limits_FC"("Settings_DB".VTD_Sys[1]);
           2:
               "Settings_DB".VTD_Sys[2] := "PopUps_DB".VTD_Settings;
               "Settings_Limits_FC"("Settings_DB".VTD_Sys[2]);
           3:
               "Settings_DB".VTD_Sys[3] := "PopUps_DB".VTD_Settings;
               "Settings_Limits_FC"("Settings_DB".VTD_Sys[3]);
           4:
               "Settings_DB".VTD_Sys[4] := "PopUps_DB".VTD_Settings;
               "Settings_Limits_FC"("Settings_DB".VTD_Sys[4]);
           5:
               "Settings_DB".VTD_Sys[5] := "PopUps_DB".VTD_Settings;
               "Settings_Limits_FC"("Settings_DB".VTD_Sys[5]);
       END_CASE;
   END_IF;

   //CONVEYORS SETTINGS
   // IF "HMI_DB".ScreenNo_Main = 10 THEN
       CASE "CNV_System_Selected" OF
           1: //SYSTEM 1
               CASE "CNV_Level_Selected" OF
                   1:
                       "Settings_DB".LCnv_Sys[1].Cnv_Level[1].Cnv1 := "PopUps_DB".Buffer_Cnv_Settings_1;
                       "Settings_DB".ECnv_Sys[1] := "PopUps_DB".ECnv_Settings;
                       "Settings_DB".LCnv_Sys[1].Cnv_Level[1].Cnv2 := "PopUps_DB".Buffer_Cnv_Settings_2;
                   2:
                       "Settings_DB".LCnv_Sys[1].Cnv_Level[2].Cnv1 := "PopUps_DB".Buffer_Cnv_Settings_1;
                       "Settings_DB".ECnv_Sys[1] := "PopUps_DB".ECnv_Settings;
                       "Settings_DB".LCnv_Sys[1].Cnv_Level[2].Cnv2 := "PopUps_DB".Buffer_Cnv_Settings_2;
                   3:
                       "Settings_DB".LCnv_Sys[1].Cnv_Level[3].Cnv1 := "PopUps_DB".Buffer_Cnv_Settings_1;
                       "Settings_DB".ECnv_Sys[1] := "PopUps_DB".ECnv_Settings;
                       "Settings_DB".LCnv_Sys[1].Cnv_Level[3].Cnv2 := "PopUps_DB".Buffer_Cnv_Settings_2;
                   4:
                       "Settings_DB".LCnv_Sys[1].Cnv_Level[4].Cnv1 := "PopUps_DB".Buffer_Cnv_Settings_1;
                       "Settings_DB".ECnv_Sys[1] := "PopUps_DB".ECnv_Settings;
                       "Settings_DB".LCnv_Sys[1].Cnv_Level[4].Cnv2 := "PopUps_DB".Buffer_Cnv_Settings_2;
                   5:
                       "Settings_DB".LCnv_Sys[1].Cnv_Level[5].Cnv1 := "PopUps_DB".Buffer_Cnv_Settings_1;
                       "Settings_DB".ECnv_Sys[1] := "PopUps_DB".ECnv_Settings;
                       "Settings_DB".LCnv_Sys[1].Cnv_Level[5].Cnv2 := "PopUps_DB".Buffer_Cnv_Settings_2;
                   6:
                       "Settings_DB".LCnv_Sys[1].Cnv_Level[6].Cnv1 := "PopUps_DB".Buffer_Cnv_Settings_1;
                       "Settings_DB".ECnv_Sys[1] := "PopUps_DB".ECnv_Settings;
                       "Settings_DB".LCnv_Sys[1].Cnv_Level[6].Cnv2 := "PopUps_DB".Buffer_Cnv_Settings_2;
                   7:
                       "Settings_DB".LCnv_Sys[1].Cnv_Level[7].Cnv1 := "PopUps_DB".Buffer_Cnv_Settings_1;
                       "Settings_DB".ECnv_Sys[1] := "PopUps_DB".ECnv_Settings;
                       "Settings_DB".LCnv_Sys[1].Cnv_Level[7].Cnv2 := "PopUps_DB".Buffer_Cnv_Settings_2;
                   8:
                       "Settings_DB".LCnv_Sys[1].Cnv_Level[8].Cnv1 := "PopUps_DB".Buffer_Cnv_Settings_1;
                       "Settings_DB".ECnv_Sys[1] := "PopUps_DB".ECnv_Settings;
                       "Settings_DB".LCnv_Sys[1].Cnv_Level[8].Cnv2 := "PopUps_DB".Buffer_Cnv_Settings_2;
               END_CASE;
           2: //SYSTEM 2
               CASE "CNV_Level_Selected" OF
                   1:
                       "Settings_DB".LCnv_Sys[2].Cnv_Level[1].Cnv1 := "PopUps_DB".Buffer_Cnv_Settings_1;
                       "Settings_DB".ECnv_Sys[2] := "PopUps_DB".ECnv_Settings;
                       "Settings_DB".LCnv_Sys[2].Cnv_Level[1].Cnv2 := "PopUps_DB".Buffer_Cnv_Settings_2;
                   2:
                       "Settings_DB".LCnv_Sys[2].Cnv_Level[2].Cnv1 := "PopUps_DB".Buffer_Cnv_Settings_1;
                       "Settings_DB".ECnv_Sys[2] := "PopUps_DB".ECnv_Settings;
                       "Settings_DB".LCnv_Sys[2].Cnv_Level[2].Cnv2 := "PopUps_DB".Buffer_Cnv_Settings_2;
                   3:
                       "Settings_DB".LCnv_Sys[2].Cnv_Level[3].Cnv1 := "PopUps_DB".Buffer_Cnv_Settings_1;
                       "Settings_DB".ECnv_Sys[2] := "PopUps_DB".ECnv_Settings;
                       "Settings_DB".LCnv_Sys[2].Cnv_Level[3].Cnv2 := "PopUps_DB".Buffer_Cnv_Settings_2;
                   4:
                       "Settings_DB".LCnv_Sys[2].Cnv_Level[4].Cnv1 := "PopUps_DB".Buffer_Cnv_Settings_1;
                       "Settings_DB".ECnv_Sys[2] := "PopUps_DB".ECnv_Settings;
                       "Settings_DB".LCnv_Sys[2].Cnv_Level[4].Cnv2 := "PopUps_DB".Buffer_Cnv_Settings_2;
                   5:
                       "Settings_DB".LCnv_Sys[2].Cnv_Level[5].Cnv1 := "PopUps_DB".Buffer_Cnv_Settings_1;
                       "Settings_DB".ECnv_Sys[2] := "PopUps_DB".ECnv_Settings;
                       "Settings_DB".LCnv_Sys[2].Cnv_Level[5].Cnv2 := "PopUps_DB".Buffer_Cnv_Settings_2;
                   6:
                       "Settings_DB".LCnv_Sys[2].Cnv_Level[6].Cnv1 := "PopUps_DB".Buffer_Cnv_Settings_1;
                       "Settings_DB".ECnv_Sys[2] := "PopUps_DB".ECnv_Settings;
                       "Settings_DB".LCnv_Sys[2].Cnv_Level[6].Cnv2 := "PopUps_DB".Buffer_Cnv_Settings_2;
                   7:
                       "Settings_DB".LCnv_Sys[2].Cnv_Level[7].Cnv1 := "PopUps_DB".Buffer_Cnv_Settings_1;
                       "Settings_DB".ECnv_Sys[2] := "PopUps_DB".ECnv_Settings;
                       "Settings_DB".LCnv_Sys[2].Cnv_Level[7].Cnv2 := "PopUps_DB".Buffer_Cnv_Settings_2;
                   8:
                       "Settings_DB".LCnv_Sys[2].Cnv_Level[8].Cnv1 := "PopUps_DB".Buffer_Cnv_Settings_1;
                       "Settings_DB".ECnv_Sys[2] := "PopUps_DB".ECnv_Settings;
                       "Settings_DB".LCnv_Sys[2].Cnv_Level[8].Cnv2 := "PopUps_DB".Buffer_Cnv_Settings_2;
               END_CASE;
           3: //SYSTEM 3
               CASE "CNV_Level_Selected" OF
                   1:
                       "Settings_DB".LCnv_Sys[3].Cnv_Level[1].Cnv1 := "PopUps_DB".Buffer_Cnv_Settings_1;
                       "Settings_DB".ECnv_Sys[3] := "PopUps_DB".ECnv_Settings;
                       "Settings_DB".LCnv_Sys[3].Cnv_Level[1].Cnv2 := "PopUps_DB".Buffer_Cnv_Settings_2;
                   2:
                       "Settings_DB".LCnv_Sys[3].Cnv_Level[2].Cnv1 := "PopUps_DB".Buffer_Cnv_Settings_1;
                       "Settings_DB".ECnv_Sys[3] := "PopUps_DB".ECnv_Settings;
                       "Settings_DB".LCnv_Sys[3].Cnv_Level[2].Cnv2 := "PopUps_DB".Buffer_Cnv_Settings_2;
                   3:
                       "Settings_DB".LCnv_Sys[3].Cnv_Level[3].Cnv1 := "PopUps_DB".Buffer_Cnv_Settings_1;
                       "Settings_DB".ECnv_Sys[3] := "PopUps_DB".ECnv_Settings;
                       "Settings_DB".LCnv_Sys[3].Cnv_Level[3].Cnv2 := "PopUps_DB".Buffer_Cnv_Settings_2;
                   4:
                       "Settings_DB".LCnv_Sys[3].Cnv_Level[4].Cnv1 := "PopUps_DB".Buffer_Cnv_Settings_1;
                       "Settings_DB".ECnv_Sys[3] := "PopUps_DB".ECnv_Settings;
                       "Settings_DB".LCnv_Sys[3].Cnv_Level[4].Cnv2 := "PopUps_DB".Buffer_Cnv_Settings_2;
                   5:
                       "Settings_DB".LCnv_Sys[3].Cnv_Level[5].Cnv1 := "PopUps_DB".Buffer_Cnv_Settings_1;
                       "Settings_DB".ECnv_Sys[3] := "PopUps_DB".ECnv_Settings;
                       "Settings_DB".LCnv_Sys[3].Cnv_Level[5].Cnv2 := "PopUps_DB".Buffer_Cnv_Settings_2;
                   6:
                       "Settings_DB".LCnv_Sys[3].Cnv_Level[6].Cnv1 := "PopUps_DB".Buffer_Cnv_Settings_1;
                       "Settings_DB".ECnv_Sys[3] := "PopUps_DB".ECnv_Settings;
                       "Settings_DB".LCnv_Sys[3].Cnv_Level[6].Cnv2 := "PopUps_DB".Buffer_Cnv_Settings_2;
                   7:
                       "Settings_DB".LCnv_Sys[3].Cnv_Level[7].Cnv1 := "PopUps_DB".Buffer_Cnv_Settings_1;
                       "Settings_DB".ECnv_Sys[3] := "PopUps_DB".ECnv_Settings;
                       "Settings_DB".LCnv_Sys[3].Cnv_Level[7].Cnv2 := "PopUps_DB".Buffer_Cnv_Settings_2;
                   8:
                       "Settings_DB".LCnv_Sys[3].Cnv_Level[8].Cnv1 := "PopUps_DB".Buffer_Cnv_Settings_1;
                       "Settings_DB".ECnv_Sys[3] := "PopUps_DB".ECnv_Settings;
                       "Settings_DB".LCnv_Sys[3].Cnv_Level[8].Cnv2 := "PopUps_DB".Buffer_Cnv_Settings_2;
               END_CASE;
           4: //SYSTEM 4
               CASE "CNV_Level_Selected" OF
                   1:
                       "Settings_DB".LCnv_Sys[4].Cnv_Level[1].Cnv1 := "PopUps_DB".Buffer_Cnv_Settings_1;
                       "Settings_DB".ECnv_Sys[4] := "PopUps_DB".ECnv_Settings;
                       "Settings_DB".LCnv_Sys[4].Cnv_Level[1].Cnv2 := "PopUps_DB".Buffer_Cnv_Settings_2;
                   2:
                       "Settings_DB".LCnv_Sys[4].Cnv_Level[2].Cnv1 := "PopUps_DB".Buffer_Cnv_Settings_1;
                       "Settings_DB".ECnv_Sys[4] := "PopUps_DB".ECnv_Settings;
                       "Settings_DB".LCnv_Sys[4].Cnv_Level[2].Cnv2 := "PopUps_DB".Buffer_Cnv_Settings_2;
                   3:
                       "Settings_DB".LCnv_Sys[4].Cnv_Level[3].Cnv1 := "PopUps_DB".Buffer_Cnv_Settings_1;
                       "Settings_DB".ECnv_Sys[4] := "PopUps_DB".ECnv_Settings;
                       "Settings_DB".LCnv_Sys[4].Cnv_Level[3].Cnv2 := "PopUps_DB".Buffer_Cnv_Settings_2;
                   4:
                       "Settings_DB".LCnv_Sys[4].Cnv_Level[4].Cnv1 := "PopUps_DB".Buffer_Cnv_Settings_1;
                       "Settings_DB".ECnv_Sys[4] := "PopUps_DB".ECnv_Settings;
                       "Settings_DB".LCnv_Sys[4].Cnv_Level[4].Cnv2 := "PopUps_DB".Buffer_Cnv_Settings_2;
                   5:
                       "Settings_DB".LCnv_Sys[4].Cnv_Level[5].Cnv1 := "PopUps_DB".Buffer_Cnv_Settings_1;
                       "Settings_DB".ECnv_Sys[4] := "PopUps_DB".ECnv_Settings;
                       "Settings_DB".LCnv_Sys[4].Cnv_Level[5].Cnv2 := "PopUps_DB".Buffer_Cnv_Settings_2;
                   6:
                       "Settings_DB".LCnv_Sys[4].Cnv_Level[6].Cnv1 := "PopUps_DB".Buffer_Cnv_Settings_1;
                       "Settings_DB".ECnv_Sys[4] := "PopUps_DB".ECnv_Settings;
                       "Settings_DB".LCnv_Sys[4].Cnv_Level[6].Cnv2 := "PopUps_DB".Buffer_Cnv_Settings_2;
                   7:
                       "Settings_DB".LCnv_Sys[4].Cnv_Level[7].Cnv1 := "PopUps_DB".Buffer_Cnv_Settings_1;
                       "Settings_DB".ECnv_Sys[4] := "PopUps_DB".ECnv_Settings;
                       "Settings_DB".LCnv_Sys[4].Cnv_Level[7].Cnv2 := "PopUps_DB".Buffer_Cnv_Settings_2;
                   8:
                       "Settings_DB".LCnv_Sys[4].Cnv_Level[8].Cnv1 := "PopUps_DB".Buffer_Cnv_Settings_1;
                       "Settings_DB".ECnv_Sys[4] := "PopUps_DB".ECnv_Settings;
                       "Settings_DB".LCnv_Sys[4].Cnv_Level[8].Cnv2 := "PopUps_DB".Buffer_Cnv_Settings_2;
               END_CASE;
           5: //SYSTEM 5
               CASE "CNV_Level_Selected" OF
                   1:
                       "Settings_DB".LCnv_Sys[5].Cnv_Level[1].Cnv1 := "PopUps_DB".Buffer_Cnv_Settings_1;
                       "Settings_DB".ECnv_Sys[5] := "PopUps_DB".ECnv_Settings;
                       "Settings_DB".LCnv_Sys[5].Cnv_Level[1].Cnv2 := "PopUps_DB".Buffer_Cnv_Settings_2;
                   2:
                       "Settings_DB".LCnv_Sys[5].Cnv_Level[2].Cnv1 := "PopUps_DB".Buffer_Cnv_Settings_1;
                       "Settings_DB".ECnv_Sys[5] := "PopUps_DB".ECnv_Settings;
                       "Settings_DB".LCnv_Sys[5].Cnv_Level[2].Cnv2 := "PopUps_DB".Buffer_Cnv_Settings_2;
                   3:
                       "Settings_DB".LCnv_Sys[5].Cnv_Level[3].Cnv1 := "PopUps_DB".Buffer_Cnv_Settings_1;
                       "Settings_DB".ECnv_Sys[5] := "PopUps_DB".ECnv_Settings;
                       "Settings_DB".LCnv_Sys[5].Cnv_Level[3].Cnv2 := "PopUps_DB".Buffer_Cnv_Settings_2;
                   4:
                       "Settings_DB".LCnv_Sys[5].Cnv_Level[4].Cnv1 := "PopUps_DB".Buffer_Cnv_Settings_1;
                       "Settings_DB".ECnv_Sys[5] := "PopUps_DB".ECnv_Settings;
                       "Settings_DB".LCnv_Sys[5].Cnv_Level[4].Cnv2 := "PopUps_DB".Buffer_Cnv_Settings_2;
                   5:
                       "Settings_DB".LCnv_Sys[5].Cnv_Level[5].Cnv1 := "PopUps_DB".Buffer_Cnv_Settings_1;
                       "Settings_DB".ECnv_Sys[5] := "PopUps_DB".ECnv_Settings;
                       "Settings_DB".LCnv_Sys[5].Cnv_Level[5].Cnv2 := "PopUps_DB".Buffer_Cnv_Settings_2;
                   6:
                       "Settings_DB".LCnv_Sys[5].Cnv_Level[6].Cnv1 := "PopUps_DB".Buffer_Cnv_Settings_1;
                       "Settings_DB".ECnv_Sys[5] := "PopUps_DB".ECnv_Settings;
                       "Settings_DB".LCnv_Sys[5].Cnv_Level[6].Cnv2 := "PopUps_DB".Buffer_Cnv_Settings_2;
                   7:
                       "Settings_DB".LCnv_Sys[5].Cnv_Level[7].Cnv1 := "PopUps_DB".Buffer_Cnv_Settings_1;
                       "Settings_DB".ECnv_Sys[5] := "PopUps_DB".ECnv_Settings;
                       "Settings_DB".LCnv_Sys[5].Cnv_Level[7].Cnv2 := "PopUps_DB".Buffer_Cnv_Settings_2;
                   8:
                       "Settings_DB".LCnv_Sys[5].Cnv_Level[8].Cnv1 := "PopUps_DB".Buffer_Cnv_Settings_1;
                       "Settings_DB".ECnv_Sys[5] := "PopUps_DB".ECnv_Settings;
                       "Settings_DB".LCnv_Sys[5].Cnv_Level[8].Cnv2 := "PopUps_DB".Buffer_Cnv_Settings_2;
               END_CASE;
       END_CASE;
   // END_IF;
END_FUNCTION

FUNCTION "PopUp_Screens_2" : Void   // FC63, SCL
{ S7_Optimized_Access := 'TRUE' }
VERSION : 0.1
// stored: AutoNumber true, IsIECCheckEnabled false, SetENOAutomatically false, UDAEnableTagReadback false
   VAR_INPUT
      HMI_No : UInt;
      HMI_Box : UInt;
      Sys_No : UInt;
   END_VAR
BEGIN
   //VTD SETTINGS
   IF "PopUps_DB_1"."VTD_Settings"[#HMI_No].ID <> 0 THEN
       "Settings_DB".VTD_Sys[#Sys_No] := "PopUps_DB_1"."VTD_Settings"[#HMI_No];
       "Settings_Limits_FC"("Settings_DB".VTD_Sys[#Sys_No]);
   END_IF;

   //CONVEYORS SETTINGS
   IF "PopUps_DB_1".ECnv_Settings[#HMI_No].ID <> 0 THEN
       CASE #HMI_Box MOD 10 OF
           1:
               "Settings_DB".LCnv_Sys[#Sys_No].Cnv_Level[1].Cnv1 := "PopUps_DB_1"."Buffer_Cnv_Settings_1"[#HMI_No];
               "Settings_DB".ECnv_Sys[#Sys_No] := "PopUps_DB_1"."ECnv_Settings"[#HMI_No];
               "Settings_DB".LCnv_Sys[#Sys_No].Cnv_Level[1].Cnv2 := "PopUps_DB_1"."Buffer_Cnv_Settings_2"[#HMI_No];
           2:
               "Settings_DB".LCnv_Sys[#Sys_No].Cnv_Level[2].Cnv1 := "PopUps_DB_1"."Buffer_Cnv_Settings_1"[#HMI_No];
               "Settings_DB".ECnv_Sys[#Sys_No] := "PopUps_DB_1"."ECnv_Settings"[#HMI_No];
               "Settings_DB".LCnv_Sys[#Sys_No].Cnv_Level[2].Cnv2 := "PopUps_DB_1"."Buffer_Cnv_Settings_2"[#HMI_No];
           3:
               "Settings_DB".LCnv_Sys[#Sys_No].Cnv_Level[3].Cnv1 := "PopUps_DB_1"."Buffer_Cnv_Settings_1"[#HMI_No];
               "Settings_DB".ECnv_Sys[#Sys_No] := "PopUps_DB_1"."ECnv_Settings"[#HMI_No];
               "Settings_DB".LCnv_Sys[#Sys_No].Cnv_Level[3].Cnv2 := "PopUps_DB_1"."Buffer_Cnv_Settings_2"[#HMI_No];
           4:
               "Settings_DB".LCnv_Sys[#Sys_No].Cnv_Level[4].Cnv1 := "PopUps_DB_1"."Buffer_Cnv_Settings_1"[#HMI_No];
               "Settings_DB".ECnv_Sys[#Sys_No] := "PopUps_DB_1"."ECnv_Settings"[#HMI_No];
               "Settings_DB".LCnv_Sys[#Sys_No].Cnv_Level[4].Cnv2 := "PopUps_DB_1"."Buffer_Cnv_Settings_2"[#HMI_No];
           5:
               "Settings_DB".LCnv_Sys[#Sys_No].Cnv_Level[5].Cnv1 := "PopUps_DB_1"."Buffer_Cnv_Settings_1"[#HMI_No];
               "Settings_DB".ECnv_Sys[#Sys_No] := "PopUps_DB_1"."ECnv_Settings"[#HMI_No];
               "Settings_DB".LCnv_Sys[#Sys_No].Cnv_Level[5].Cnv2 := "PopUps_DB_1"."Buffer_Cnv_Settings_2"[#HMI_No];
           6:
               "Settings_DB".LCnv_Sys[#Sys_No].Cnv_Level[6].Cnv1 := "PopUps_DB_1"."Buffer_Cnv_Settings_1"[#HMI_No];
               "Settings_DB".ECnv_Sys[#Sys_No] := "PopUps_DB_1"."ECnv_Settings"[#HMI_No];
               "Settings_DB".LCnv_Sys[#Sys_No].Cnv_Level[6].Cnv2 := "PopUps_DB_1"."Buffer_Cnv_Settings_2"[#HMI_No];
           7:
               "Settings_DB".LCnv_Sys[#Sys_No].Cnv_Level[7].Cnv1 := "PopUps_DB_1"."Buffer_Cnv_Settings_1"[#HMI_No];
               "Settings_DB".ECnv_Sys[#Sys_No] := "PopUps_DB_1"."ECnv_Settings"[#HMI_No];
               "Settings_DB".LCnv_Sys[#Sys_No].Cnv_Level[7].Cnv2 := "PopUps_DB_1"."Buffer_Cnv_Settings_2"[#HMI_No];
           8:
               "Settings_DB".LCnv_Sys[#Sys_No].Cnv_Level[8].Cnv1 := "PopUps_DB_1"."Buffer_Cnv_Settings_1"[#HMI_No];
               "Settings_DB".ECnv_Sys[#Sys_No] := "PopUps_DB_1"."ECnv_Settings"[#HMI_No];
               "Settings_DB".LCnv_Sys[#Sys_No].Cnv_Level[8].Cnv2 := "PopUps_DB_1"."Buffer_Cnv_Settings_2"[#HMI_No];
       END_CASE;
   END_IF;
END_FUNCTION

FUNCTION "Post_Safe" : Void   // FC1001, LAD
{ S7_Optimized_Access := 'TRUE' }
VERSION : 0.1
// stored: AutoNumber false, IsIECCheckEnabled false, SetENOAutomatically false, UDAEnableTagReadback false
BEGIN

REGION Network 1
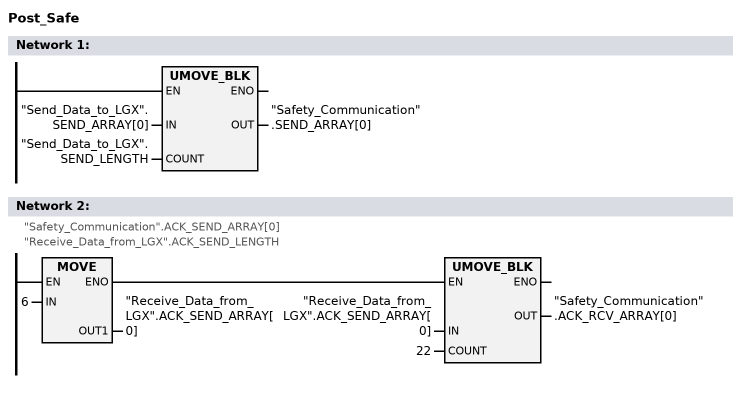
   UMOVE_BLK(IN := "Send_Data_to_LGX".SEND_ARRAY[0],
             COUNT := "Send_Data_to_LGX".SEND_LENGTH,
             OUT => "Safety_Communication".SEND_ARRAY[0]);
END_REGION

REGION Network 2
   // "Safety_Communication".ACK_SEND_ARRAY[0]
   // 
   // 
   // "Receive_Data_from_LGX".ACK_SEND_LENGTH
   "Receive_Data_from_LGX".ACK_SEND_ARRAY[0] := 6;
   UMOVE_BLK(IN := "Receive_Data_from_LGX".ACK_SEND_ARRAY[0],
             COUNT := 22,
             OUT => "Safety_Communication".ACK_RCV_ARRAY[0]);
END_REGION
END_FUNCTION

FUNCTION "Pre_Safe" : Void   // FC1000, LAD
{ S7_Optimized_Access := 'TRUE' }
VERSION : 0.1
// stored: AutoNumber false, IsIECCheckEnabled false, SetENOAutomatically false, UDAEnableTagReadback false
BEGIN

REGION Network 1
   // "Receive_Data_from_LGX".RCV_LENGTH
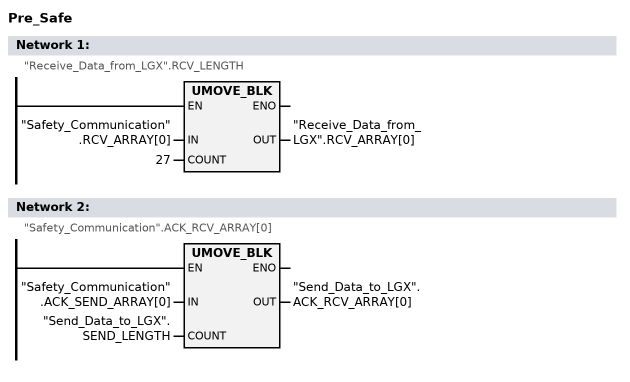
   UMOVE_BLK(IN := "Safety_Communication".RCV_ARRAY[0],
             COUNT := 27,
             OUT => "Receive_Data_from_LGX".RCV_ARRAY[0]);
END_REGION

REGION Network 2
   // "Safety_Communication".ACK_RCV_ARRAY[0]
   UMOVE_BLK(IN := "Safety_Communication".ACK_SEND_ARRAY[0],
             COUNT := "Send_Data_to_LGX".SEND_LENGTH,
             OUT => "Send_Data_to_LGX".ACK_RCV_ARRAY[0]);
END_REGION
END_FUNCTION

FUNCTION "RemovePlusSign" : String   // FC14, SCL
{ S7_Optimized_Access := 'TRUE' }
VERSION : 0.1
// stored: AutoNumber true, IsIECCheckEnabled false, SetENOAutomatically false, UDAEnableTagReadback false
   VAR_INPUT
      inString : String;
   END_VAR
   VAR_TEMP
      tempString : String;
   END_VAR
BEGIN

   IF LEFT(IN := #inString, L := 1) = '+' THEN
       #tempString := RIGHT(IN := #inString, L := LEN(#inString) - 1);
   ELSE
       #tempString := #inString;
   END_IF;

   #RemovePlusSign := #tempString;
END_FUNCTION

FUNCTION "SICK_GetValue" : Void   // FC10, SCL
TITLE = Get value
{ S7_Optimized_Access := 'TRUE' }
AUTHOR : SICKAG
FAMILY : Ident
VERSION : 1.0
// This function is needs to get a value out of a SICK CoLa command.
// stored: AutoNumber false, IsIECCheckEnabled false, SetENOAutomatically false, UDAEnableTagReadback false
   VAR_INPUT
      iTelegramLength : UInt;   // Length of the source telegram
      iValueLength : USInt;   // ASCII length of the value [1..8] = Fix length | [0]= Variable
      arrData : Array[0..499] of Byte;   // Data record (contains the whole CoLa telegram)
   END_VAR
   VAR_OUTPUT
      nValue : DWord;   // Read value
      nErrorCode : Word;   // Error code
   END_VAR
   VAR_IN_OUT
      iPosition : UInt;   // Position offset of the value before and after (starting from 0)
   END_VAR
   VAR_TEMP
      iLoop : Int;   // Temporarily variable
      iSegmentLength : UInt;   // Length of the segement
      nTemp : DWord;   // Temporarily variable
   END_VAR
BEGIN
   (*===========================================================================================
   Name:   SICK_GetValue
   Author: SICK AG
   =============================================================================================
   Description: 
   This function is for internal use only. The function gets the selected Hex-value string out 
   of the CoLa-Telegram and convert it into a hexadecimal number. 

   =============================================================================================
   Error codes:
   16#0000 = No error
   16#0001 = Invaild telegram length   
   16#0002 = Invalid position index 
   16#0003 = Invalid value length
   16#0004 = Invalid segment length 
   16#0005 = ASCII character is not in a hexadecimal format             

   =============================================================================================
   Version history:
   Date       | Version | created under               | Author  | Remark
   ---------------------------------------------------------------------------------------------
   30/01/2014 | V1.0    | TIA Portal V12 SP1 Update 2 | SICK AG | Initial version
   ============================================================================================*)

   (*===================================== INITIALISATION =====================================*)
   #iSegmentLength:= 0;
   #nValue:= 16#0000_0000;
   #nErrorCode:= 16#0000;

   (*======================================= READ VALUE =======================================*)
   (*Check telegram length*)
   IF #iTelegramLength <=0 OR #iTelegramLength > 500 THEN
     #nErrorCode:= 16#0001; (*Error: Invaild telegram length*)
     RETURN;
   END_IF;

   (*Check current position of the value*)
   IF #iPosition > (#iTelegramLength-1) THEN
     #nErrorCode:= 16#0002; (*Error: Invalid position index*)
     RETURN;
   END_IF;

   (*Check value length*)
   IF #iValueLength >8 THEN
     #nErrorCode:= 16#0003; (*Error: Invalid value length*)
     RETURN;
   END_IF;

   (*Get a value with a variable length (ends with a ' ' or [ETX]*)
   IF #iValueLength = 0 THEN
     FOR #iLoop:= UINT_TO_INT(#iPosition) TO UINT_TO_INT(#iTelegramLength-1) DO
       (*Check if a blank or a [ETX] is detected*)
       IF (#arrData[#iLoop] =' ') OR (#arrData[#iLoop] ='$03') THEN
         EXIT;
       END_IF;

       (*Length of the current value segement*)
       #iSegmentLength:= #iSegmentLength+1;
     END_FOR;

   (*Get a value with a fixed character length [1..8]*)
   ELSE
     #iSegmentLength:= #iValueLength;
   END_IF;

   (*Check if the segment length is valid*)
   IF (#iSegmentLength >8) OR (#iSegmentLength =0) THEN
     #nErrorCode:= 16#0004; (*Error: Invalid segment length*)
     RETURN;
   END_IF;

   (*Convert ASCII string into a hexadecimal number*)
   FOR #iLoop:= UINT_TO_INT(#iPosition) TO UINT_TO_INT(#iPosition+#iSegmentLength-1) DO
     (*ACSII value = [0..9]*)
     IF #arrData[#iLoop] >='0' AND #arrData[#iLoop] <='9' THEN
       #nTemp:= #arrData[#iLoop]-48;
     (*ASCII value = [A..F]*) 
     ELSIF #arrData[#iLoop] >='A' AND #arrData[#iLoop] <='F' THEN
       #nTemp:= #arrData[#iLoop]-55;
     (*ASCII value = [a..f]*)
     ELSIF #arrData[#iLoop] >='a' AND #arrData[#iLoop] <='f' THEN
       #nTemp:= #arrData[#iLoop]-87;    
     ELSE
       #nErrorCode:= 16#0005; (*Error: ASCII character is not in a hexadecimal format *)
       RETURN;
     END_IF;

     (*Create hexadecimal number*)
     #nValue:= SHL(IN:= #nValue, N:= 4);
     #nValue:= #nValue+#nTemp;
   END_FOR;

   (*Set the position of the next element in the telegram*)
   IF #iValueLength = 0 THEN
     #iPosition:= #iPosition+#iSegmentLength+1; (*With blank character*)
   ELSE
     #iPosition:= #iPosition+#iSegmentLength; (*Without blank character*)
   END_IF;
END_FUNCTION

FUNCTION "SICK_SetValue" : Void   // FC11, SCL
TITLE = Set value
{ S7_Optimized_Access := 'TRUE' }
AUTHOR : SICKAG
FAMILY : Ident
VERSION : 1.1
// This function is needs to set a value to a SICK CoLa command.
// stored: AutoNumber false, IsIECCheckEnabled false, SetENOAutomatically false, UDAEnableTagReadback false
   VAR_INPUT
      bAddBlank : Bool;   // Add blank after value
      nValue : DWord;   // Value that should be written
   END_VAR
   VAR_OUTPUT
      arrData : Array[0..499] of Byte;   // Destination telegram
      nErrorCode : Word;   // Error code
   END_VAR
   VAR_IN_OUT
      iPosition : UInt;   // Position offset of the value before and after (starting from 0)
   END_VAR
   VAR_TEMP
      iValueLength : USInt;   // Byte length of the value that shuld be written
      nReturnValue : Word;   // Return value of the convert function
      sValue : String[8];   // Converted value
      nTempValue : DWord;   // Temporarily variable
      iTemp : UInt;   // Temporarily variable
   END_VAR
BEGIN
   (*===========================================================================================
   Name:   SICK_SetValue
   Author: SICK AG
   =============================================================================================
   Description: 
   This function is for internal use only.
   The function converts a hexadecimal value into a hexadecimal string and add it 
   automatically to the command array.     

   =============================================================================================
   Error codes:
   16#0000 = No error
   16#0001 = Invalid position index   
   16#8xxx = Conversion error (HTA-Function) see help system for more information

   =============================================================================================
   Version history:
   Date       | Version | created under               | Author  | Remark
   ---------------------------------------------------------------------------------------------
   30/01/2014 | V1.0    | TIA Portal V12 SP1 Update 2 | SICK AG | Initial version
   22/04/2014 | V1.1    | TIA Portal V12 SP1 Update 4 | SICK AG | Avoid warnings that occur with 
                                                                  TIA V13
   ============================================================================================*)

   (*===================================== INITIALISATION =====================================*)
   #iValueLength:= 0;
   #nErrorCode:= 16#0000;

   (*======================================= WRITE VALUE ======================================*)
   (*Check current position of the value*)
   IF #iPosition > 499 THEN 
     #nErrorCode:= 16#0001; (*Error: Invalid position index*)
     RETURN;
   END_IF;



   (*Get byte length of the value that should be written*)
   IF #nValue <= 16#FF THEN
     #nTempValue:= SHL(IN:= #nValue, N:=24);
     #iValueLength:= 1;
   ELSIF #nValue <= 16#FFFF THEN
     #nTempValue:= SHL(IN:= #nValue, N:=16);
     #iValueLength:= 2;
   ELSIF #nValue <= 16#00FF_FFFF THEN
     #nTempValue:= SHL(IN:= #nValue, N:=8);
     #iValueLength:= 3;
   ELSIF #nValue <= 16#FFFF_FFFF THEN
     #nTempValue:= #nValue;
     #iValueLength:= 4;
   END_IF;

   (*Convert hexadecimal number into a ASCII string*)
   #nReturnValue:= HTA(IN:= #nTempValue, N:= #iValueLength, OUT=>#sValue);
   IF #nReturnValue <> 16#0000 THEN
     #nErrorCode:= #nReturnValue; (*Error: Conversion error (HTA-Function)*)
     RETURN;
   END_IF;

   (*Add the string value to the destination telegram*)
   #arrData[#iPosition]:= 0; // Avoid warnings under TIA V13
   Strg_TO_Chars(Strg:=#sValue, pChars:= #iPosition, Cnt=> #iTemp, Chars:= #arrData);

   (*Add blank to the destination telegram and calculate the position of the next element*)
   IF #bAddBlank THEN
     #arrData[#iPosition+#iTemp]:= ' ';
     #iPosition:= #iPosition+#iTemp+1;

   (*Calculate the position of the next element*)
   ELSE
     #iPosition:= #iPosition+#iTemp;
   END_IF;
END_FUNCTION

FUNCTION "Safety_Data_FC" : Void   // FC50, SCL
{ S7_Optimized_Access := 'TRUE' }
VERSION : 0.1
// stored: AutoNumber true, IsIECCheckEnabled false, SetENOAutomatically false, UDAEnableTagReadback false
   VAR_INPUT
      C1101_EStop : Bool;
      C1102_EStop : Bool;
      C1103_EStop : Bool;
      C1101_LG1 : Bool;
      C1101_LG2 : Bool;
      C1102_LG1 : Bool;
      C1102_LG2 : Bool;
      C1103_LG1 : Bool;
      C1103_LG2 : Bool;
   END_VAR
   VAR_OUTPUT
      o_LGX_Zone01_EStop : Bool;
      o_LGX_Zone02_EStop : Bool;
      o_LGX_Zone03_EStop : Bool;
      o_LGX_Zone04_EStop : Bool;
      o_LGX_Zone05_EStop : Bool;
      o_LGX_Zone06_EStop : Bool;
      o_LGX_Zone07_EStop : Bool;
      o_LGX_Zone08_EStop : Bool;
      o_LGX_Zone09_EStop : Bool;
      o_LGX_Zone10_EStop : Bool;
      o_LGX_Infeed_I1103_CS : Bool;
      o_LGX_Infeed_I1105_CS : Bool;
      o_LGX_Infeed_I1107_CS : Bool;
      o_LGX_Outfeed_I1401_CS : Bool;
      o_LGX_Outfeed_I1403_CS : Bool;
      o_LGX_Outfeed_I1407_CS : Bool;
      o_Any_LGX_EStop_Active : Bool;
      o_Any_LGX_Conv_CS_Active : Bool;
   END_VAR
BEGIN
   // // ============================================================
   // // FC_Safety_PreProcess (FC1000 on the Spacemaker side)
   // // Safety data pre-processing before OPC-UA transmission
   // // Execute in the F-Runtime Group (Main_Safety_RTG1)
   // // Ref: Section 6 of the document
   // // ============================================================

   // // NOTE: This FC runs in the F-Runtime safety group (Safety Program).
   // // Inputs are the actual safety signals from the SM system.
   // // Outputs populate the safety DB that will be published by the OPC-UA Server.

   // // --- Map E-Stops to SM → LGX safety DB ---
   // "DB_Safety_SM_To_LGX".VTD_I1310_EStop_Active := #C1101_EStop;
   // "DB_Safety_SM_To_LGX".VTD_I1320_EStop_Active := #C1102_EStop;
   // "DB_Safety_SM_To_LGX".VTD_I1330_EStop_Active := #C1103_EStop;

   // // --- Map Light Guards ---
   // "DB_Safety_SM_To_LGX".VTD_I1310_LG1_Active := #C1101_LG1;
   // "DB_Safety_SM_To_LGX".VTD_I1310_LG2_Active := #C1101_LG2;
   // "DB_Safety_SM_To_LGX".VTD_I1320_LG1_Active := #C1102_LG1;
   // "DB_Safety_SM_To_LGX".VTD_I1320_LG2_Active := #C1102_LG2;
   // "DB_Safety_SM_To_LGX".VTD_I1330_LG1_Active := #C1103_LG1;
   // "DB_Safety_SM_To_LGX".VTD_I1330_LG2_Active := #C1103_LG2;


   // // ============================================================
   // // FC_Safety_PostProcess (FC1001 on the Spacemaker side)
   // // Post-processing of safety data received from LGX
   // // Execute in the F-Runtime Group (Main_Safety_RTG1)
   // // Ref: Section 6 of the document
   // // ============================================================

   // // --- Map received data from LGX DB → SM Safety ---
   // #o_LGX_Zone01_EStop := "DB_Safety_LGX_To_SM".Zone_01_EStop_Active;
   // #o_LGX_Zone02_EStop := "DB_Safety_LGX_To_SM".Zone_02_EStop_Active;
   // #o_LGX_Zone03_EStop := "DB_Safety_LGX_To_SM".Zone_03_EStop_Active;
   // #o_LGX_Zone04_EStop := "DB_Safety_LGX_To_SM".Zone_04_EStop_Active;
   // #o_LGX_Zone05_EStop := "DB_Safety_LGX_To_SM".Zone_05_EStop_Active;
   // #o_LGX_Zone06_EStop := "DB_Safety_LGX_To_SM".Zone_06_EStop_Active;
   // #o_LGX_Zone07_EStop := "DB_Safety_LGX_To_SM".Zone_07_EStop_Active;
   // #o_LGX_Zone08_EStop := "DB_Safety_LGX_To_SM".Zone_08_EStop_Active;
   // #o_LGX_Zone09_EStop := "DB_Safety_LGX_To_SM".Zone_09_EStop_Active;
   // #o_LGX_Zone10_EStop := "DB_Safety_LGX_To_SM".Zone_10_EStop_Active;

   // #o_LGX_Infeed_I1103_CS := "DB_Safety_LGX_To_SM".Infeed_I1103_CS;
   // #o_LGX_Infeed_I1105_CS := "DB_Safety_LGX_To_SM".Infeed_I1105_CS;
   // #o_LGX_Infeed_I1107_CS := "DB_Safety_LGX_To_SM".Infeed_I1107_CS;

   // #o_LGX_Outfeed_I1401_CS := "DB_Safety_LGX_To_SM".Outfeed_I1401_CS;
   // #o_LGX_Outfeed_I1403_CS := "DB_Safety_LGX_To_SM".Outfeed_I1403_CS;
   // #o_LGX_Outfeed_I1407_CS := "DB_Safety_LGX_To_SM".Outfeed_I1407_CS;

   // // --- Consolidated flags for use in SM safety logic ---
   // #o_Any_LGX_EStop_Active :=
   // #o_LGX_Zone01_EStop OR #o_LGX_Zone02_EStop OR #o_LGX_Zone03_EStop OR
   // #o_LGX_Zone04_EStop OR #o_LGX_Zone05_EStop OR #o_LGX_Zone06_EStop OR
   // #o_LGX_Zone07_EStop OR #o_LGX_Zone08_EStop OR #o_LGX_Zone09_EStop OR
   // #o_LGX_Zone10_EStop;

   // #o_Any_LGX_Conv_CS_Active :=
   // #o_LGX_Infeed_I1103_CS OR #o_LGX_Infeed_I1105_CS OR #o_LGX_Infeed_I1107_CS OR
   // #o_LGX_Outfeed_I1401_CS OR #o_LGX_Outfeed_I1403_CS OR #o_LGX_Outfeed_I1407_CS;
END_FUNCTION

FUNCTION "Screens" : Void   // FC12, SCL
{ S7_Optimized_Access := 'TRUE' }
VERSION : 0.1
// stored: AutoNumber true, IsIECCheckEnabled false, SetENOAutomatically false, UDAEnableTagReadback false
   VAR_TEMP
      i : UInt;
      j : UInt;
      _id_decoded_OP : Array[1..5] of "ID_Decoded";
      Level_Strg : String;
      Destination_Location : Array[1..5] of DInt;
   END_VAR
BEGIN
   REGION MAIN SCREEN
       REGION AUTOMATIC BUTTON - SYSTEM 1
           IF "Automatic_Button_1" THEN
               FOR #i := "Settings_DB".VTD_Sys[1].Lowest_Level TO "Settings_DB".VTD_Sys[1].Highest_Level DO
                   "Control_DB".VTD_Sys[1].Instruction.Mode_Change :=
                   "Control_DB".ECnv_Sys[1].Instruction.Mode_Change :=
                   "Control_DB".LCnv_Sys[1].Cnv_Level[#i].Cnv1.Instruction.Mode_Change :=
                   "Control_DB".LCnv_Sys[1].Cnv_Level[#i].Cnv2.Instruction.Mode_Change :=
                   "Control_DB".LCnv_Sys[1].Cnv_Level[#i].Cnv1.Safety_Stop_Cnrl.Mode :=
                   "Control_DB".LCnv_Sys[1].Cnv_Level[#i].Cnv2.Safety_Stop_Cnrl.Mode := 3;

                   "Control_DB".VTD_Sys[1].Instruction.Enable :=
                   "Control_DB".ECnv_Sys[1].Instruction.Enable :=
                   "Control_DB".LCnv_Sys[1].Cnv_Level[#i].Cnv1.Instruction.Enable :=
                   "Control_DB".LCnv_Sys[1].Cnv_Level[#i].Cnv2.Instruction.Enable := TRUE;
               END_FOR;
           END_IF;
       END_REGION

       REGION AUTOMATIC BUTTON - SYSTEM 2
           IF "Automatic_Button_2" THEN
               FOR #i := "Settings_DB".VTD_Sys[2].Lowest_Level TO "Settings_DB".VTD_Sys[2].Highest_Level DO
                   "Control_DB".VTD_Sys[2].Instruction.Mode_Change :=
                   "Control_DB".ECnv_Sys[2].Instruction.Mode_Change :=
                   "Control_DB".LCnv_Sys[2].Cnv_Level[#i].Cnv1.Instruction.Mode_Change :=
                   "Control_DB".LCnv_Sys[2].Cnv_Level[#i].Cnv2.Instruction.Mode_Change :=
                   "Control_DB".LCnv_Sys[2].Cnv_Level[#i].Cnv1.Safety_Stop_Cnrl.Mode :=
                   "Control_DB".LCnv_Sys[2].Cnv_Level[#i].Cnv2.Safety_Stop_Cnrl.Mode := 3;

                   "Control_DB".VTD_Sys[2].Instruction.Enable :=
                   "Control_DB".ECnv_Sys[2].Instruction.Enable :=
                   "Control_DB".LCnv_Sys[2].Cnv_Level[#i].Cnv1.Instruction.Enable :=
                   "Control_DB".LCnv_Sys[2].Cnv_Level[#i].Cnv2.Instruction.Enable := TRUE;
               END_FOR;
           END_IF;
       END_REGION

       REGION AUTOMATIC BUTTON - SYSTEM 3
           IF "Automatic_Button_3" THEN
               FOR #i := "Settings_DB".VTD_Sys[3].Lowest_Level TO "Settings_DB".VTD_Sys[3].Highest_Level DO
                   "Control_DB".VTD_Sys[3].Instruction.Mode_Change :=
                   "Control_DB".ECnv_Sys[3].Instruction.Mode_Change :=
                   "Control_DB".LCnv_Sys[3].Cnv_Level[#i].Cnv1.Instruction.Mode_Change :=
                   "Control_DB".LCnv_Sys[3].Cnv_Level[#i].Cnv2.Instruction.Mode_Change :=
                   "Control_DB".LCnv_Sys[3].Cnv_Level[#i].Cnv1.Safety_Stop_Cnrl.Mode :=
                   "Control_DB".LCnv_Sys[3].Cnv_Level[#i].Cnv2.Safety_Stop_Cnrl.Mode := 3;

                   "Control_DB".VTD_Sys[3].Instruction.Enable :=
                   "Control_DB".ECnv_Sys[3].Instruction.Enable :=
                   "Control_DB".LCnv_Sys[3].Cnv_Level[#i].Cnv1.Instruction.Enable :=
                   "Control_DB".LCnv_Sys[3].Cnv_Level[#i].Cnv2.Instruction.Enable := TRUE;
               END_FOR;
           END_IF;
       END_REGION

       REGION AUTOMATIC BUTTON - SYSTEM 4
           IF "Automatic_Button_4" THEN
               FOR #i := "Settings_DB".VTD_Sys[4].Lowest_Level TO "Settings_DB".VTD_Sys[4].Highest_Level DO
                   "Control_DB".VTD_Sys[4].Instruction.Mode_Change :=
                   "Control_DB".ECnv_Sys[4].Instruction.Mode_Change :=
                   "Control_DB".LCnv_Sys[4].Cnv_Level[#i].Cnv1.Instruction.Mode_Change :=
                   "Control_DB".LCnv_Sys[4].Cnv_Level[#i].Cnv2.Instruction.Mode_Change :=
                   "Control_DB".LCnv_Sys[4].Cnv_Level[#i].Cnv1.Safety_Stop_Cnrl.Mode :=
                   "Control_DB".LCnv_Sys[4].Cnv_Level[#i].Cnv2.Safety_Stop_Cnrl.Mode := 3;

                   "Control_DB".VTD_Sys[4].Instruction.Enable :=
                   "Control_DB".ECnv_Sys[4].Instruction.Enable :=
                   "Control_DB".LCnv_Sys[4].Cnv_Level[#i].Cnv1.Instruction.Enable :=
                   "Control_DB".LCnv_Sys[4].Cnv_Level[#i].Cnv2.Instruction.Enable := TRUE;
               END_FOR;
           END_IF;
       END_REGION

       REGION AUTOMATIC BUTTON - SYSTEM 5
           IF "Automatic_Button_5" THEN
               FOR #i := "Settings_DB".VTD_Sys[5].Lowest_Level TO "Settings_DB".VTD_Sys[5].Highest_Level DO
                   "Control_DB".VTD_Sys[5].Instruction.Mode_Change :=
                   "Control_DB".ECnv_Sys[5].Instruction.Mode_Change :=
                   "Control_DB".LCnv_Sys[5].Cnv_Level[#i].Cnv1.Instruction.Mode_Change :=
                   "Control_DB".LCnv_Sys[5].Cnv_Level[#i].Cnv2.Instruction.Mode_Change :=
                   "Control_DB".LCnv_Sys[5].Cnv_Level[#i].Cnv1.Safety_Stop_Cnrl.Mode :=
                   "Control_DB".LCnv_Sys[5].Cnv_Level[#i].Cnv2.Safety_Stop_Cnrl.Mode := 3;

                   "Control_DB".VTD_Sys[5].Instruction.Enable :=
                   "Control_DB".ECnv_Sys[5].Instruction.Enable :=
                   "Control_DB".LCnv_Sys[5].Cnv_Level[#i].Cnv1.Instruction.Enable :=
                   "Control_DB".LCnv_Sys[5].Cnv_Level[#i].Cnv2.Instruction.Enable := TRUE;
               END_FOR;
           END_IF;
       END_REGION

       REGION ALL IN AUTOMATIC - SYSTEM 1
           "All_In_Automatic_1" := "Control_DB".VTD_Sys[1].Mode = 3 AND //VTD
           "Control_DB".ECnv_Sys[1].Mode = 3 AND //ECONVEYOR
           //CONVEYORS
           "Control_DB".LCnv_Sys[1].Cnv_Level[1].Cnv1.Mode = 3 AND
           "Control_DB".LCnv_Sys[1].Cnv_Level[1].Cnv2.Mode = 3 AND
           "Control_DB".LCnv_Sys[1].Cnv_Level[2].Cnv1.Mode = 3 AND
           "Control_DB".LCnv_Sys[1].Cnv_Level[2].Cnv2.Mode = 3 AND
           "Control_DB".LCnv_Sys[1].Cnv_Level[3].Cnv1.Mode = 3 AND
           "Control_DB".LCnv_Sys[1].Cnv_Level[3].Cnv2.Mode = 3 AND
           "Control_DB".LCnv_Sys[1].Cnv_Level[4].Cnv1.Mode = 3 AND
           "Control_DB".LCnv_Sys[1].Cnv_Level[4].Cnv2.Mode = 3 AND
           "Control_DB".LCnv_Sys[1].Cnv_Level[5].Cnv1.Mode = 3 AND
           "Control_DB".LCnv_Sys[1].Cnv_Level[5].Cnv2.Mode = 3 AND
           "Control_DB".LCnv_Sys[1].Cnv_Level[6].Cnv1.Mode = 3 AND
           "Control_DB".LCnv_Sys[1].Cnv_Level[6].Cnv2.Mode = 3 AND
           "Control_DB".LCnv_Sys[1].Cnv_Level[7].Cnv1.Mode = 3 AND
           "Control_DB".LCnv_Sys[1].Cnv_Level[7].Cnv2.Mode = 3 AND
           "Control_DB".LCnv_Sys[1].Cnv_Level[8].Cnv1.Mode = 3 AND
           "Control_DB".LCnv_Sys[1].Cnv_Level[8].Cnv2.Mode = 3 AND
           //SAFETY STOP
           "Control_DB".LCnv_Sys[1].Cnv_Level[1].Cnv1.Safety_Stop_Cnrl.Mode = 3 AND
           "Control_DB".LCnv_Sys[1].Cnv_Level[1].Cnv2.Safety_Stop_Cnrl.Mode = 3 AND
           "Control_DB".LCnv_Sys[1].Cnv_Level[2].Cnv1.Safety_Stop_Cnrl.Mode = 3 AND
           "Control_DB".LCnv_Sys[1].Cnv_Level[2].Cnv2.Safety_Stop_Cnrl.Mode = 3 AND
           "Control_DB".LCnv_Sys[1].Cnv_Level[3].Cnv1.Safety_Stop_Cnrl.Mode = 3 AND
           "Control_DB".LCnv_Sys[1].Cnv_Level[3].Cnv2.Safety_Stop_Cnrl.Mode = 3 AND
           "Control_DB".LCnv_Sys[1].Cnv_Level[4].Cnv1.Safety_Stop_Cnrl.Mode = 3 AND
           "Control_DB".LCnv_Sys[1].Cnv_Level[4].Cnv2.Safety_Stop_Cnrl.Mode = 3 AND
           "Control_DB".LCnv_Sys[1].Cnv_Level[5].Cnv1.Safety_Stop_Cnrl.Mode = 3 AND
           "Control_DB".LCnv_Sys[1].Cnv_Level[5].Cnv2.Safety_Stop_Cnrl.Mode = 3 AND
           "Control_DB".LCnv_Sys[1].Cnv_Level[6].Cnv1.Safety_Stop_Cnrl.Mode = 3 AND
           "Control_DB".LCnv_Sys[1].Cnv_Level[6].Cnv2.Safety_Stop_Cnrl.Mode = 3 AND
           "Control_DB".LCnv_Sys[1].Cnv_Level[7].Cnv1.Safety_Stop_Cnrl.Mode = 3 AND
           "Control_DB".LCnv_Sys[1].Cnv_Level[7].Cnv2.Safety_Stop_Cnrl.Mode = 3 AND
           "Control_DB".LCnv_Sys[1].Cnv_Level[8].Cnv1.Safety_Stop_Cnrl.Mode = 3 AND
           "Control_DB".LCnv_Sys[1].Cnv_Level[8].Cnv2.Safety_Stop_Cnrl.Mode = 3;
       END_REGION

       REGION ALL IN AUTOMATIC - SYSTEM 2
           "All_In_Automatic_2" := "Control_DB".VTD_Sys[2].Mode = 3 AND //VTD
           "Control_DB".ECnv_Sys[2].Mode = 3 AND //ECONVEYOR
           //CONVEYORS
           "Control_DB".LCnv_Sys[2].Cnv_Level[1].Cnv1.Mode = 3 AND
           "Control_DB".LCnv_Sys[2].Cnv_Level[1].Cnv2.Mode = 3 AND
           "Control_DB".LCnv_Sys[2].Cnv_Level[2].Cnv1.Mode = 3 AND
           "Control_DB".LCnv_Sys[2].Cnv_Level[2].Cnv2.Mode = 3 AND
           "Control_DB".LCnv_Sys[2].Cnv_Level[3].Cnv1.Mode = 3 AND
           "Control_DB".LCnv_Sys[2].Cnv_Level[3].Cnv2.Mode = 3 AND
           "Control_DB".LCnv_Sys[2].Cnv_Level[4].Cnv1.Mode = 3 AND
           "Control_DB".LCnv_Sys[2].Cnv_Level[4].Cnv2.Mode = 3 AND
           "Control_DB".LCnv_Sys[2].Cnv_Level[5].Cnv1.Mode = 3 AND
           "Control_DB".LCnv_Sys[2].Cnv_Level[5].Cnv2.Mode = 3 AND
           "Control_DB".LCnv_Sys[2].Cnv_Level[6].Cnv1.Mode = 3 AND
           "Control_DB".LCnv_Sys[2].Cnv_Level[6].Cnv2.Mode = 3 AND
           "Control_DB".LCnv_Sys[2].Cnv_Level[7].Cnv1.Mode = 3 AND
           "Control_DB".LCnv_Sys[2].Cnv_Level[7].Cnv2.Mode = 3 AND
           "Control_DB".LCnv_Sys[2].Cnv_Level[8].Cnv1.Mode = 3 AND
           "Control_DB".LCnv_Sys[2].Cnv_Level[8].Cnv2.Mode = 3 AND
           //SAFETY STOP
           "Control_DB".LCnv_Sys[2].Cnv_Level[1].Cnv1.Safety_Stop_Cnrl.Mode = 3 AND
           "Control_DB".LCnv_Sys[2].Cnv_Level[1].Cnv2.Safety_Stop_Cnrl.Mode = 3 AND
           "Control_DB".LCnv_Sys[2].Cnv_Level[2].Cnv1.Safety_Stop_Cnrl.Mode = 3 AND
           "Control_DB".LCnv_Sys[2].Cnv_Level[2].Cnv2.Safety_Stop_Cnrl.Mode = 3 AND
           "Control_DB".LCnv_Sys[2].Cnv_Level[3].Cnv1.Safety_Stop_Cnrl.Mode = 3 AND
           "Control_DB".LCnv_Sys[2].Cnv_Level[3].Cnv2.Safety_Stop_Cnrl.Mode = 3 AND
           "Control_DB".LCnv_Sys[2].Cnv_Level[4].Cnv1.Safety_Stop_Cnrl.Mode = 3 AND
           "Control_DB".LCnv_Sys[2].Cnv_Level[4].Cnv2.Safety_Stop_Cnrl.Mode = 3 AND
           "Control_DB".LCnv_Sys[2].Cnv_Level[5].Cnv1.Safety_Stop_Cnrl.Mode = 3 AND
           "Control_DB".LCnv_Sys[2].Cnv_Level[5].Cnv2.Safety_Stop_Cnrl.Mode = 3 AND
           "Control_DB".LCnv_Sys[2].Cnv_Level[6].Cnv1.Safety_Stop_Cnrl.Mode = 3 AND
           "Control_DB".LCnv_Sys[2].Cnv_Level[6].Cnv2.Safety_Stop_Cnrl.Mode = 3 AND
           "Control_DB".LCnv_Sys[2].Cnv_Level[7].Cnv1.Safety_Stop_Cnrl.Mode = 3 AND
           "Control_DB".LCnv_Sys[2].Cnv_Level[7].Cnv2.Safety_Stop_Cnrl.Mode = 3 AND
           "Control_DB".LCnv_Sys[2].Cnv_Level[8].Cnv1.Safety_Stop_Cnrl.Mode = 3 AND
           "Control_DB".LCnv_Sys[2].Cnv_Level[8].Cnv2.Safety_Stop_Cnrl.Mode = 3;
       END_REGION

       REGION ALL IN AUTOMATIC - SYSTEM 3
           "All_In_Automatic_3" := "Control_DB".VTD_Sys[3].Mode = 3 AND //VTD
           "Control_DB".ECnv_Sys[3].Mode = 3 AND //ECONVEYOR
           //CONVEYORS
           "Control_DB".LCnv_Sys[3].Cnv_Level[1].Cnv1.Mode = 3 AND
           "Control_DB".LCnv_Sys[3].Cnv_Level[1].Cnv2.Mode = 3 AND
           "Control_DB".LCnv_Sys[3].Cnv_Level[2].Cnv1.Mode = 3 AND
           "Control_DB".LCnv_Sys[3].Cnv_Level[2].Cnv2.Mode = 3 AND
           "Control_DB".LCnv_Sys[3].Cnv_Level[3].Cnv1.Mode = 3 AND
           "Control_DB".LCnv_Sys[3].Cnv_Level[3].Cnv2.Mode = 3 AND
           "Control_DB".LCnv_Sys[3].Cnv_Level[4].Cnv1.Mode = 3 AND
           "Control_DB".LCnv_Sys[3].Cnv_Level[4].Cnv2.Mode = 3 AND
           "Control_DB".LCnv_Sys[3].Cnv_Level[5].Cnv1.Mode = 3 AND
           "Control_DB".LCnv_Sys[3].Cnv_Level[5].Cnv2.Mode = 3 AND
           "Control_DB".LCnv_Sys[3].Cnv_Level[6].Cnv1.Mode = 3 AND
           "Control_DB".LCnv_Sys[3].Cnv_Level[6].Cnv2.Mode = 3 AND
           "Control_DB".LCnv_Sys[3].Cnv_Level[7].Cnv1.Mode = 3 AND
           "Control_DB".LCnv_Sys[3].Cnv_Level[7].Cnv2.Mode = 3 AND
           "Control_DB".LCnv_Sys[3].Cnv_Level[8].Cnv1.Mode = 3 AND
           "Control_DB".LCnv_Sys[3].Cnv_Level[8].Cnv2.Mode = 3 AND
           //SAFETY STOP
           "Control_DB".LCnv_Sys[3].Cnv_Level[1].Cnv1.Safety_Stop_Cnrl.Mode = 3 AND
           "Control_DB".LCnv_Sys[3].Cnv_Level[1].Cnv2.Safety_Stop_Cnrl.Mode = 3 AND
           "Control_DB".LCnv_Sys[3].Cnv_Level[2].Cnv1.Safety_Stop_Cnrl.Mode = 3 AND
           "Control_DB".LCnv_Sys[3].Cnv_Level[2].Cnv2.Safety_Stop_Cnrl.Mode = 3 AND
           "Control_DB".LCnv_Sys[3].Cnv_Level[3].Cnv1.Safety_Stop_Cnrl.Mode = 3 AND
           "Control_DB".LCnv_Sys[3].Cnv_Level[3].Cnv2.Safety_Stop_Cnrl.Mode = 3 AND
           "Control_DB".LCnv_Sys[3].Cnv_Level[4].Cnv1.Safety_Stop_Cnrl.Mode = 3 AND
           "Control_DB".LCnv_Sys[3].Cnv_Level[4].Cnv2.Safety_Stop_Cnrl.Mode = 3 AND
           "Control_DB".LCnv_Sys[3].Cnv_Level[5].Cnv1.Safety_Stop_Cnrl.Mode = 3 AND
           "Control_DB".LCnv_Sys[3].Cnv_Level[5].Cnv2.Safety_Stop_Cnrl.Mode = 3 AND
           "Control_DB".LCnv_Sys[3].Cnv_Level[6].Cnv1.Safety_Stop_Cnrl.Mode = 3 AND
           "Control_DB".LCnv_Sys[3].Cnv_Level[6].Cnv2.Safety_Stop_Cnrl.Mode = 3 AND
           "Control_DB".LCnv_Sys[3].Cnv_Level[7].Cnv1.Safety_Stop_Cnrl.Mode = 3 AND
           "Control_DB".LCnv_Sys[3].Cnv_Level[7].Cnv2.Safety_Stop_Cnrl.Mode = 3 AND
           "Control_DB".LCnv_Sys[3].Cnv_Level[8].Cnv1.Safety_Stop_Cnrl.Mode = 3 AND
           "Control_DB".LCnv_Sys[3].Cnv_Level[8].Cnv2.Safety_Stop_Cnrl.Mode = 3;
       END_REGION

       REGION ALL IN AUTOMATIC - SYSTEM 4
           "All_In_Automatic_4" := "Control_DB".VTD_Sys[4].Mode = 3 AND //VTD
           "Control_DB".ECnv_Sys[4].Mode = 3 AND //ECONVEYOR
           //CONVEYORS
           "Control_DB".LCnv_Sys[4].Cnv_Level[1].Cnv1.Mode = 3 AND
           "Control_DB".LCnv_Sys[4].Cnv_Level[2].Cnv1.Mode = 3 AND
           "Control_DB".LCnv_Sys[4].Cnv_Level[3].Cnv1.Mode = 3 AND
           "Control_DB".LCnv_Sys[4].Cnv_Level[4].Cnv1.Mode = 3 AND
           "Control_DB".LCnv_Sys[4].Cnv_Level[5].Cnv1.Mode = 3 AND
           "Control_DB".LCnv_Sys[4].Cnv_Level[6].Cnv1.Mode = 3 AND
           "Control_DB".LCnv_Sys[4].Cnv_Level[7].Cnv1.Mode = 3 AND
           "Control_DB".LCnv_Sys[4].Cnv_Level[8].Cnv1.Mode = 3 AND
           //SAFETY STOP
           "Control_DB".LCnv_Sys[4].Cnv_Level[1].Cnv1.Safety_Stop_Cnrl.Mode = 3 AND
           "Control_DB".LCnv_Sys[4].Cnv_Level[2].Cnv1.Safety_Stop_Cnrl.Mode = 3 AND
           "Control_DB".LCnv_Sys[4].Cnv_Level[3].Cnv1.Safety_Stop_Cnrl.Mode = 3 AND
           "Control_DB".LCnv_Sys[4].Cnv_Level[4].Cnv1.Safety_Stop_Cnrl.Mode = 3 AND
           "Control_DB".LCnv_Sys[4].Cnv_Level[5].Cnv1.Safety_Stop_Cnrl.Mode = 3 AND
           "Control_DB".LCnv_Sys[4].Cnv_Level[6].Cnv1.Safety_Stop_Cnrl.Mode = 3 AND
           "Control_DB".LCnv_Sys[4].Cnv_Level[7].Cnv1.Safety_Stop_Cnrl.Mode = 3 AND
           "Control_DB".LCnv_Sys[4].Cnv_Level[8].Cnv1.Safety_Stop_Cnrl.Mode = 3;
       END_REGION

       REGION ALL IN AUTOMATIC - SYSTEM 5
           "All_In_Automatic_5" := "Control_DB".VTD_Sys[5].Mode = 3 AND //VTD
           "Control_DB".ECnv_Sys[5].Mode = 3 AND //ECONVEYOR
           //CONVEYORS
           "Control_DB".LCnv_Sys[5].Cnv_Level[1].Cnv1.Mode = 3 AND
           "Control_DB".LCnv_Sys[5].Cnv_Level[2].Cnv1.Mode = 3 AND
           "Control_DB".LCnv_Sys[5].Cnv_Level[3].Cnv1.Mode = 3 AND
           "Control_DB".LCnv_Sys[5].Cnv_Level[4].Cnv1.Mode = 3 AND
           "Control_DB".LCnv_Sys[5].Cnv_Level[5].Cnv1.Mode = 3 AND
           "Control_DB".LCnv_Sys[5].Cnv_Level[6].Cnv1.Mode = 3 AND
           "Control_DB".LCnv_Sys[5].Cnv_Level[7].Cnv1.Mode = 3 AND
           "Control_DB".LCnv_Sys[5].Cnv_Level[8].Cnv1.Mode = 3 AND
           //SAFETY STOP
           "Control_DB".LCnv_Sys[5].Cnv_Level[1].Cnv1.Safety_Stop_Cnrl.Mode = 3 AND
           "Control_DB".LCnv_Sys[5].Cnv_Level[2].Cnv1.Safety_Stop_Cnrl.Mode = 3 AND
           "Control_DB".LCnv_Sys[5].Cnv_Level[3].Cnv1.Safety_Stop_Cnrl.Mode = 3 AND
           "Control_DB".LCnv_Sys[5].Cnv_Level[4].Cnv1.Safety_Stop_Cnrl.Mode = 3 AND
           "Control_DB".LCnv_Sys[5].Cnv_Level[5].Cnv1.Safety_Stop_Cnrl.Mode = 3 AND
           "Control_DB".LCnv_Sys[5].Cnv_Level[6].Cnv1.Safety_Stop_Cnrl.Mode = 3 AND
           "Control_DB".LCnv_Sys[5].Cnv_Level[7].Cnv1.Safety_Stop_Cnrl.Mode = 3 AND
           "Control_DB".LCnv_Sys[5].Cnv_Level[8].Cnv1.Safety_Stop_Cnrl.Mode = 3;
       END_REGION

       "Bypass".Main_Panel.ACK := "Reset_Comissioning";

       REGION Order processing
           //DECODES
           #Destination_Location[1] := "System_DB_1".OrderTable[1].OPC_Control.Destination_Location;
           #Destination_Location[2] := "System_DB_2".OrderTable[1].OPC_Control.Destination_Location;
           #Destination_Location[3] := "System_DB_3".OrderTable[1].OPC_Control.Destination_Location;
           #Destination_Location[4] := "System_DB_4".OrderTable[1].OPC_Control.Destination_Location;
           #Destination_Location[5] := "System_DB_5".OrderTable[1].OPC_Control.Destination_Location;

           FOR #i := 1 TO "Settings_DB".System.VTD_Count DO
               "ID_Decode_F"(ID := #Destination_Location[#i],
                             ID_Decoded := #_id_decoded_OP[#i]);
           END_FOR;

           //CLASSIFIES
           FOR #i := 1 TO "Settings_DB".System.VTD_Count DO
               IF #_id_decoded_OP[#i].Level <> 0 THEN
                   VAL_STRG(IN := #_id_decoded_OP[#i].Level,
                            FORMAT := 16#0000,
                            PREC := 0,
                            P := 1,
                            SIZE := 0,
                            OUT => #Level_Strg);
                   CASE #_id_decoded_OP[#i].VTD OF
                       1: //System 1
                           IF #_id_decoded_OP[#i].Device_Type = 30 THEN //VTD
                               "Screen_DB".OrderProcessing[#i] := CONCAT(IN1 := "System_DB_1".OrderTable[1].Device, IN2 := ' To LEVEL ', IN3 := #Level_Strg);
                           ELSIF #_id_decoded_OP[#i].Device_Type = 10 THEN //CNV1
                               "Screen_DB".OrderProcessing[#i] := CONCAT(IN1 := "System_DB_1".OrderTable[1].Device, IN2 := ' To CNV 1 LEVEL ', IN3 := #Level_Strg);
                           ELSIF #_id_decoded_OP[#i].Device_Type = 11 THEN //CNV2
                               "Screen_DB".OrderProcessing[#i] := CONCAT(IN1 := "System_DB_1".OrderTable[1].Device, IN2 := ' To CNV 2 LEVEL ', IN3 := #Level_Strg);
                           ELSIF #_id_decoded_OP[#i].Device_Type = 12 THEN //ECONVEYOR
                               "Screen_DB".OrderProcessing[#i] := CONCAT(IN1 := "System_DB_1".OrderTable[1].Device, IN2 := ' To ECONV LEVEL ', IN3 := #Level_Strg);
                           END_IF;

                       2: //System 2
                           IF #_id_decoded_OP[#i].Device_Type = 30 THEN //VTD
                               "Screen_DB".OrderProcessing[#i] := CONCAT(IN1 := "System_DB_2".OrderTable[1].Device, IN2 := ' To LEVEL ', IN3 := #Level_Strg);
                           ELSIF #_id_decoded_OP[#i].Device_Type = 10 THEN //CNV1
                               "Screen_DB".OrderProcessing[#i] := CONCAT(IN1 := "System_DB_2".OrderTable[1].Device, IN2 := ' To CNV 1 LEVEL ', IN3 := #Level_Strg);
                           ELSIF #_id_decoded_OP[#i].Device_Type = 11 THEN //CNV2
                               "Screen_DB".OrderProcessing[#i] := CONCAT(IN1 := "System_DB_2".OrderTable[1].Device, IN2 := ' To CNV 2 LEVEL ', IN3 := #Level_Strg);
                           ELSIF #_id_decoded_OP[#i].Device_Type = 12 THEN //ECONVEYOR
                               "Screen_DB".OrderProcessing[#i] := CONCAT(IN1 := "System_DB_2".OrderTable[1].Device, IN2 := ' To ECONV LEVEL ', IN3 := #Level_Strg);
                           END_IF;

